(* IEC 61131-3 sources: brOscatLib/oscatBasic (part 3) *)

(* ---- REVERSE.st ---- *)
FUNCTION REVERSE
    (*http://www.oscat.de/images/OSCATBasic/oscat_basic333_en.pdf#page=232*)
    (* new code donated by rebler wolfgang *)
    REVERSE := ROR(IN,1) AND 2#10001000 OR ROL(IN,1) AND 2#00010001 OR ROR(IN,3) AND 2#01000100 OR ROL(IN,3) AND 2#00100010;

    (* old code
    REVERSE := SHL(IN,7) OR SHR(IN,7) OR (ROR(IN,3) AND 2#01000100) OR (ROL(IN,3) AND 2#00100010)
    	OR (SHL(IN,1) AND 2#00010000) OR (SHR(IN,1) AND 2#00001000);
    *)

    (* revision history
    hm		9.oct 2007		rev 1.0
    	original version

    hm		18. feb 2008	rev 1.1
    	improved performance

    RW    3. feb. 2021  	rev 1.2
    	improved performance
    *)
END_FUNCTION

(* ---- RND.st ---- *)
FUNCTION RND
    (*http://www.oscat.de/images/OSCATBasic/oscat_basic333_en.pdf#page=64*)
    IF X = 0.0 THEN
    	RND := 0.0;
    ELSE
    	M := EXPN(10.0,N - CEIL(LOG(ABS(X))));
    	RND := DINT_TO_REAL(REAL_TO_DINT(X * M)) / M;
    END_IF

    (* revision history
    hm	11. mar 2008	rev 1.0
    	original version

    hm	26. oct. 2008	rev 1.1
    	code optimization

    hm	10. mar. 2009	rev 1.2
    	real constants updated to new systax using dot

    *)

END_FUNCTION

(* ---- ROUND.st ---- *)
FUNCTION ROUND
    (*http://www.oscat.de/images/OSCATBasic/oscat_basic333_en.pdf#page=65*)
    X := cDECADES[LIMIT(0,N,8)];
    ROUND := DINT_TO_REAL(REAL_TO_DINT(IN * X)) / X;

    (* revision history
    hm	1. sep 2006	rev 1.0
    	original version

    hm	2. dec 2007	rev 1.1
    	changed code for better performance

    hm	8. jan 2008	rev 1.2
    	further improvement IN performance

    hm 11. mar. 2008	rev 1.3
    	corrected an error with negative numbers
    	use real_to_dint instead of trunc

    hm	16. mar 2008	rev 1.4
    	added type conversion to avoid warning under codesys 3.0

    hm	25. oct. 2008	rev 1.5
    	new code using global constants decades
    *)

END_FUNCTION

(* ---- SCALE.st ---- *)
FUNCTION SCALE
    (*http://www.oscat.de/images/OSCATBasic/oscat_basic333_en.pdf#page=288*)
    SCALE := LIMIT(MN, X * K + O, MX);

    (* revision history
    hm	16. may. 2008		rev 1.0
    	original version
    *)
END_FUNCTION

(* ---- SCALE_B.st ---- *)
FUNCTION SCALE_B
    (*http://www.oscat.de/images/OSCATBasic/oscat_basic333_en.pdf#page=289*)
    _I_HI := BYTE_TO_USINT(I_HI);
    _I_LO := BYTE_TO_USINT(I_LO);
    IF I_HI = I_LO THEN
    	SCALE_B := O_LO;
    ELSE
    	SCALE_B := (O_HI - O_LO) / USINT_TO_REAL(_I_HI - _I_LO) * USINT_TO_REAL(LIMIT(_I_LO, BYTE_TO_USINT(X), _I_HI));
    END_IF

    (* revision history
    hm	18. may. 2008		rev 1.0
    	original version

    hm	18. jan 2011		rev 1.1
    	avoid division by 0

    *)
END_FUNCTION

(* ---- SCALE_B2.st ---- *)
FUNCTION SCALE_B2
    (*http://www.oscat.de/images/OSCATBasic/oscat_basic333_en.pdf#page=290*)
    SCALE_B2 := 	(((IN1_MAX - IN1_MIN)* BYTE_TO_USINT(IN1) + (IN2_MAX - IN2_MIN)* BYTE_TO_USINT(IN2)) * 0.003921569 + IN1_MIN + IN2_MIN) * K + O;

    (* revision History
    hm 19.1.2007		rev 1.1
    	changed outputs to real to avoid overflow of integer
    	added offset for better cascading of scale functions
    	changed from FB to function

    hm	6. jan 2008		rev 1.2
    	improved performance

    hm	26. oct. 2008	rev 1.3
    	code optimization

    hm	3. nov. 2008	rev 1.4
    	used wrong factor in formula

    *)
END_FUNCTION

(* ---- SCALE_B4.st ---- *)
FUNCTION SCALE_B4
    (*http://www.oscat.de/images/OSCATBasic/oscat_basic333_en.pdf#page=291*)
    SCALE_B4 := 	(((IN1_MAX - IN1_MIN)* BYTE_TO_USINT(IN1) + (IN2_MAX - IN2_MIN)* BYTE_TO_USINT(IN2) + (IN3_MAX - IN3_MIN)* BYTE_TO_USINT(IN3) + (IN4_MAX - IN4_MIN)* BYTE_TO_USINT(IN4))* 0.003921569 + IN1_MIN + IN2_MIN + IN3_MIN + IN4_MIN) * K + O;

    (* revision History
    hm 19.1.2007		rev 1.1
    	changed outputs to real to avoid overflow of integer
    	added offset for better cascading of scale functions
    	changed from fb to function

    hm	6. jan 2008		rev 1.2
    	improved performance

    hm	26. oct. 2008	rev 1.3
    	optimized code

    hm	3. nov. 2008	rev 1.4
    	used wrong factor in formula

    *)
END_FUNCTION

(* ---- SCALE_B8.st ---- *)
FUNCTION SCALE_B8
    (*http://www.oscat.de/images/OSCATBasic/oscat_basic333_en.pdf#page=292*)
    SCALE_B8 := 	(((IN1_MAX - IN1_MIN)* BYTE_TO_USINT(IN1) + (IN2_MAX - IN2_MIN)* BYTE_TO_USINT(IN2) + (IN3_MAX - IN3_MIN)* BYTE_TO_USINT(IN3) + (IN4_MAX - IN4_MIN)* BYTE_TO_USINT(IN4) +
    				(IN5_MAX - IN5_MIN)* BYTE_TO_USINT(IN5) + (IN6_MAX - IN6_MIN)* BYTE_TO_USINT(IN6) + (IN7_MAX - IN7_MIN)* BYTE_TO_USINT(IN7) + (IN8_MAX - IN8_MIN)* BYTE_TO_USINT(IN8)) * 0.003921569
    				 + IN1_MIN + IN2_MIN + IN3_MIN + IN4_MIN + IN5_MIN + IN6_MIN + IN7_MIN + IN8_MIN) * K + O;

    (* revision History
    hm	19. jan.2007	rev 1.1
    	changed outputs to real to avoid overflow of integer
    	added offset for better cascading of scale functions

    hm	6. jan. 2008	rev 1.2
    	improved performance

    hm	26. oct. 2008	rev 1.3
    	code optimization

    hm	3. nov. 2008	rev 1.4
    	used wrong factor in formula

    *)
END_FUNCTION

(* ---- SCALE_D.st ---- *)
FUNCTION SCALE_D
    (*http://www.oscat.de/images/OSCATBasic/oscat_basic333_en.pdf#page=293*)
    _I_HI := DWORD_TO_UDINT(I_HI);
    _I_LO := DWORD_TO_UDINT(I_LO);
    IF _I_HI = _I_LO THEN
    	SCALE_D := O_LO;
    ELSE
    	SCALE_D := (O_HI - O_LO) / UDINT_TO_REAL(_I_HI - _I_LO) * UDINT_TO_REAL(LIMIT(_I_LO, DWORD_TO_UDINT(X), _I_HI) - _I_LO) + O_LO;
    END_IF

    (* revision history
    hm	18. may. 2008	rev 1.0
    	original version

    hm	13. nov. 2008	rev 1.1
    	corrected formula for negative gradient

    hm	11. jan 2011	rev 1.2
    	avoid division by 0
    *)
END_FUNCTION

(* ---- SCALE_R.st ---- *)
FUNCTION SCALE_R
    (*http://www.oscat.de/images/OSCATBasic/oscat_basic333_en.pdf#page=294*)
    IF I_LO = I_HI THEN
    	SCALE_R := O_LO;
    ELSE
    	SCALE_R := (O_HI - O_LO) / (I_HI - I_LO) * (LIMIT(I_LO, X, I_HI) - I_LO) + O_LO;
    END_IF

    (* revision history
    hm	18. may. 2008	rev 1.0
    	original version

    hm	13. nov. 2008	rev 1.1
    	corrected formula for negative gradient

    hm	11. jan 2011	rev 1.2
    	avoid division by 0

    *)
END_FUNCTION

(* ---- SCALE_X2.st ---- *)
FUNCTION SCALE_X2
    (*http://www.oscat.de/images/OSCATBasic/oscat_basic333_en.pdf#page=295*)
    SCALE_X2 := (SEL(IN1, IN1_MIN, IN1_MAX)+ SEL(IN2, IN2_MIN, IN2_MAX)) * K + O;

    (* revision history
    hm	19. jan, 2007	rev 1.0
    	original version

    hm	26. oct. 2008	rev 1.1
    	code optimized

    *)
END_FUNCTION

(* ---- SCALE_X4.st ---- *)
FUNCTION SCALE_X4
    (*http://www.oscat.de/images/OSCATBasic/oscat_basic333_en.pdf#page=296*)
    SCALE_X4 := (SEL(IN1,IN1_MIN, IN1_MAX) + SEL(IN2, IN2_MIN, IN2_MAX)+SEL(IN3, IN3_MIN, IN3_MAX)+ SEL(IN4, IN4_MIN, IN4_MAX)) * K + O;

    (* revision history
    hm	19. jan. 2008	rev 1.0
    	original version

    hm	26. oct. 2008	rev 1.1
    	optimized code
    *)
END_FUNCTION

(* ---- SCALE_X8.st ---- *)
FUNCTION SCALE_X8
    (*http://www.oscat.de/images/OSCATBasic/oscat_basic333_en.pdf#page=297*)
    SCALE_X8 := (SEL(IN1,IN1_MIN, IN1_MAX)+ SEL(IN2,IN2_MIN, IN2_MAX)+SEL(IN3,IN3_MIN, IN3_MAX)+ SEL(IN4,IN4_MIN, IN4_MAX)
    				+SEL(IN5,IN5_MIN, IN5_MAX)+ SEL(IN6,IN6_MIN, IN6_MAX)+SEL(IN7,IN7_MIN, IN7_MAX)+ SEL(IN8,IN8_MIN, IN8_MAX)) * K + O;

    (* revision history
    hm	19. jan. 2008	rev 1.0
    	original version

    hm	26. oct. 2008	rev 1.1
    	optimized code

    hm	24. jan. 2008	rev 1.2
    	corrected error in formula
    *)
END_FUNCTION

(* ---- SDT_TO_DATE.st ---- *)
FUNCTION SDT_TO_DATE
    (*http://www.oscat.de/images/OSCATBasic/oscat_basic333_en.pdf#page=134*)
    SDT_TO_DATE := SET_DATE(DTI.YEAR, DTI.MONTH, DTI.DAY);

    (* revision history

    hm 18. oct. 2008	rev 1.0
    	original version

    *)
END_FUNCTION

(* ---- SDT_TO_DT.st ---- *)
FUNCTION SDT_TO_DT
    (*http://www.oscat.de/images/OSCATBasic/oscat_basic333_en.pdf#page=135*)
    SDT_TO_DT := SET_DT(DTI.YEAR, DTI.MONTH, DTI.DAY, DTI.HOUR, DTI.MINUTE, DTI.SECOND);

    (* revision history

    hm 18. oct. 2008	rev 1.0
    	original version

    *)
END_FUNCTION

(* ---- SDT_TO_TOD.st ---- *)
FUNCTION SDT_TO_TOD
    (*http://www.oscat.de/images/OSCATBasic/oscat_basic333_en.pdf#page=135*)
    SDT_TO_TOD := UDINT_TO_TOD(INT_TO_UDINT(DTI.HOUR) * 3600000 + INT_TO_UDINT(DTI.MINUTE) * 60000 + INT_TO_UDINT(DTI.SECOND) * 1000 + INT_TO_UDINT(DTI.MS));

    (* revision history

    hm 18. oct. 2008	rev 1.0
    	original version

    hm	16. nov. 2008	rev 1.1
    	added typecasts to avoid warnings
    *)
END_FUNCTION

(* ---- SECOND.st ---- *)
FUNCTION SECOND
    (*http://www.oscat.de/images/OSCATBasic/oscat_basic333_en.pdf#page=135*)
    SECOND := UDINT_TO_REAL(TOD_TO_UDINT(ITOD) - TOD_TO_UDINT(ITOD)/60000 * 60000) / 1000.0;

    (* change history

    hm	2. oct. 2006 rev 1.1
    	changed name of input to ITOD

    *)
END_FUNCTION

(* ---- SECOND_OF_DT.st ---- *)
FUNCTION SECOND_OF_DT
    (*http://www.oscat.de/images/OSCATBasic/oscat_basic333_en.pdf#page=136*)
    SECOND_OF_DT := UDINT_TO_INT(DT_TO_UDINT(XDT) MOD 60);

    (* revision history
    hm		6.9.2008	rev 1.0
    	original version

    *)
END_FUNCTION

(* ---- SECOND_TO_TIME.st ---- *)
FUNCTION SECOND_TO_TIME
    (*http://www.oscat.de/images/OSCATBasic/oscat_basic333_en.pdf#page=136*)
    SECOND_TO_TIME := DWORD_TO_TIME(REAL_TO_DWORD(IN * 1000.0));

    (* revision history
    hm	4. aug. 2006	rev 1.0
    	original version

    hm	14. mar. 2008	rev 1.1
    	rounded the input after the last digit

    hm	24. feb. 2009	rev 1.2
    	changed input to IN
    *)
END_FUNCTION

(* ---- SENSOR_INT.st ---- *)
FUNCTION SENSOR_INT
    (*http://www.oscat.de/images/OSCATBasic/oscat_basic333_en.pdf#page=324*)
    IF CURRENT <> 0.0 THEN
    	RG := VOLTAGE / CURRENT;
    	SENSOR_INT := RP * ( RG - RS) / ( RP + RS - RG);
    END_IF

    (* revisaion history

    hm 20.1.2007		rev 1.1
    	deleted input R0 which was not needed.

    hm	2. dec 2007	rev 1.2
    	corrected an error in formula and improoved speed

    hm	11. mar. 2009	rev 1.3
    	changed real constants to use dot syntax

    *)
END_FUNCTION

(* ---- SET_DATE.st ---- *)
FUNCTION SET_DATE
    (*http://www.oscat.de/images/OSCATBasic/oscat_basic333_en.pdf#page=136*)
    IF (MONTH > 2) AND (SHL(YEAR,14) = 0)
    THEN (* we add one DAY for leap YEAR *)
    	SET_DATE := UDINT_TO_DATE((INT_TO_UDINT(ofs[MONTH] + DAY ) + SHR(INT_TO_UDINT(YEAR) * 1461 - 2878169, 2))*86400);
    ELSE
    	SET_DATE := UDINT_TO_DATE((INT_TO_UDINT(ofs[MONTH] + DAY - 1 ) + SHR(INT_TO_UDINT(YEAR) * 1461 - 2878169, 2))*86400);
    END_IF

    (* old code
    IF MONTH > 2 THEN
    	count := (MONTH - 1) * 30;
    	IF MONTH > 7 THEN count := count + SHR(MONTH - 3,1); ELSE count := count + SHR(MONTH - 4,1); END_IF
    	(* chech for leap YEAR and add one DAY if true
    	IF SHL(YEAR,14) = 0 THEN count := count + 1; END_IF
    ELSE
    	count := (MONTH - 1) * 31;
    END_IF

    SET_DATE := UDINT_TO_DATE((INT_TO_UDINT(count + DAY - 1) + SHR(INT_TO_UDINT(YEAR) * 1461 - 2878169, 2)) * 86400);
    *)

    (* revision history
    hm	4. aug. 2006	rev 1.0
    	original version

    hm	19 sep. 2007	rev 1.1
    	use function leap_year to calculate leap YEAR, more exceptions are handled

    hm	1. okt	2007	rev 1.2
    	added compatibility to step7

    hm	16.dec 2007		rev 1.3
    	changed code to improove performance

    hm	3. jan. 2008	rev 1.4
    	further improvements in performance

    hm	16. mar. 2008	rev 1.5
    	added type conversions to avoid warnings under codesys 3.0

    hm	7. apr. 2008	rev 1.6
    	deleted unused step7 code

    hm	14. oct. 2008	rev 1.7
    	optimized code for better performance

    hm	25. oct. 2008	rev 2.0
    	new code using setup constants

    hm	16. nov. 2008	rev 2.1
    	added typecasts to avoid warnings

    hm	22. jan. 2011	rev 2.2
    	improved performance

    hm	29. dec. 2011	rev 2.3
    	improved performance

    hm 3. FEB 2021 rev 2.4
    	new code to be more readable
    *)
END_FUNCTION

(* ---- SET_DT.st ---- *)
FUNCTION SET_DT
    (*http://www.oscat.de/images/OSCATBasic/oscat_basic333_en.pdf#page=137*)
    SET_DT := UDINT_TO_DT(DATE_TO_UDINT(SET_DATE(YEAR, MONTH, DAY)) + INT_TO_UDINT(SECOND) + INT_TO_UDINT(MINUTE) * 60 + INT_TO_UDINT(HOUR) * 3600);

    (* revision history
    hm	4. aug. 2006		rev 1.0
    	original version

    hm		19 sep. 2007	rev 1.1
    	use function leap_year to calculate leap YEAR, more exceptions are handled

    hm		1. okt 2007		rev 1.2
    	added step7 compatibility
    	call function set_date

    hm		8. oct 2007		rev 1.3
    	deleted unused variables count and leap

    hm		1. 11 2007		rev 1.4
    	converted HOUR type integer to dword in calculation to avoid overrun on möller ecp4

    hm		16. mar 2008	rev 1.5
    	added type conversions to avoid warnings under codesys 3.0
    *)

END_FUNCTION

(* ---- SET_TOD.st ---- *)
FUNCTION SET_TOD
    (*http://www.oscat.de/images/OSCATBasic/oscat_basic333_en.pdf#page=138*)
    SET_TOD := UDINT_TO_TOD(REAL_TO_UDINT(SECOND * 1000.0) + INT_TO_UDINT(MINUTE) * 60000 + INT_TO_UDINT(HOUR) * 3600000);

    (* revision history

    hm		4.aug.2006		rev 1.0
    	original version

    hm		11. sep 2007	rev 1.1
    	changed coding to avoid a compiler warning under twincat.

    hm		1. nov 2007	rev 1.2
    	changed coding to avoid possible overrun situation on möller ecp4

    hm		2. Nov	2007	rev 1.3
    	changed dword to DINT in calcualtion to avoid warnings with some compilers

    hm		14. mar 2008	rev 1.4
    	changed code to avoid rounding problem at last digit of millisecond

    hm		16. mar. 2008	rev 1.5
    	added type conversions to avoid warning under codesys 3.0
    *)
END_FUNCTION

(* ---- SGN.st ---- *)
FUNCTION SGN
    (*http://www.oscat.de/images/OSCATBasic/oscat_basic333_en.pdf#page=65*)
    IF X > 0 THEN
    	SGN := 1;
    ELSIF X < 0 THEN
    	SGN := -1;
    ELSE
    	SGN := 0;
    END_IF

    (* revision histroy
    hm	16. oct 2007	rev 1.0
    	original version

    hm	11. nov 2007	rev 1.1
    	changed type of function from real to int

    *)
END_FUNCTION

(* ---- SHL1.st ---- *)
FUNCTION SHL1
    (*http://www.oscat.de/images/OSCATBasic/oscat_basic333_en.pdf#page=233*)
    SHL1 := SHR(temp,32-N) OR SHL(IN,N);

    (* revision history
    hm	14.9.2007		rev 1.0
    	original version

    hm	27. dec 2007	rev 1.1
    	changed code for better performance

    *)
END_FUNCTION

(* ---- SHR1.st ---- *)
FUNCTION SHR1
    (*http://www.oscat.de/images/OSCATBasic/oscat_basic333_en.pdf#page=233*)
    SHR1 := SHL(temp,32-N) OR SHR(IN,N);

    (* revision history
    hm	14.9.2007		rev 1.0
    	original version

    hm	27. dec 2007	rev 1.1
    	changed code for better performance

    *)
END_FUNCTION

(* ---- SIGMOID.st ---- *)
FUNCTION SIGMOID
    (*http://www.oscat.de/images/OSCATBasic/oscat_basic333_en.pdf#page=66*)
    IF X > 20.0 THEN
    	SIGMOID := 1.0;
    ELSIF X < -85.0 THEN
    	SIGMOID := 0.0;
    ELSE
    	SIGMOID := 1.0 / (1.0 + EXP(-X));
    END_IF

    (* revision history
    hm	10.12.2007		rev 1.0
    	original version

    hm	11. mar. 2008		rev 1.1
    	extended range of valid inputs to +inv / -inv

    hm 10. mar. 2009		rev 1.2
    	real constants updated to new systax using dot

    *)
END_FUNCTION

(* ---- SIGN_I.st ---- *)
FUNCTION SIGN_I
    (*http://www.oscat.de/images/OSCATBasic/oscat_basic333_en.pdf#page=66*)
    SIGN_I := IN.31;

    (* revision history
    hm 3.3.2007	rev 1.1
    	changed method of function for better compatibility to other systems

    hm	1.12.2007	rev 1.2
    	changed code to improve performance

    hm	27. oct. 2008	rev 1.3
    	changed type of input to dint

    *)
END_FUNCTION

(* ---- SIGN_R.st ---- *)
FUNCTION SIGN_R
    (*http://www.oscat.de/images/OSCATBasic/oscat_basic333_en.pdf#page=67*)
    SIGN_R := IN < 0.0;

    (* revision history
    hm 19.1.2007	rev 1.1
    	changed method of function for better compatibility to other systems

    hm	1.12.2007	rev 1.2
    	changed code to improve performance

    hm	14. jun. 2008	rev 1.3
    	improved performace

    hm 10. mar. 2009	rev 1.4
    	real constants updated to new systax using dot

    *)
END_FUNCTION

(* ---- SINC.st ---- *)
FUNCTION SINC
    (*http://www.oscat.de/images/OSCATBasic/oscat_basic333_en.pdf#page=67*)
    IF X = 0.0 THEN
    	SINC := 1.0;
    ELSE
    	SINC := SIN(X) / X;
    END_IF

    (* revision histroy
    hm	11. mar. 2008	rev 1.0
    	original version

    hm	1.12.2007	rev 1.1
    	changed code to improove performance

    hm 10. mar. 2009	rev 1.2
    	real constants updated to new systax using dot

    *)
END_FUNCTION

(* ---- SINH.st ---- *)
FUNCTION SINH
    (*http://www.oscat.de/images/OSCATBasic/oscat_basic333_en.pdf#page=67*)
    IF ABS(X) < 2E-3 THEN
    	SINH := X;
    ELSE
    	SINH := (EXP(X) - EXP(-X)) * 0.5;
    END_IF

    (* revision history
    hm	12.1.2007	rev 1.0
    	original version

    hm	1.12.2007	rev 1.1
    	changed code to improve performance

    hm	5. jan 2008	rev 1.2
    	further performance improvement

    hm	11. mar 2008	rev 1.3
    	improved accuracy around 0

    *)
END_FUNCTION

(* ---- SPHERE_V.st ---- *)
FUNCTION SPHERE_V
    (*http://www.oscat.de/images/OSCATBasic/oscat_basic333_en.pdf#page=106*)
    SPHERE_V := 4.188790205 * RX * RX * RX;

    (* revision histroy
    hm	16. oct 2007	rev 1.0
    	original version

    hm	4. dec 2007		rev 1.1
    	changed code for better performance

    hm	22. feb 2008		rev 1.2
    	changed code for better performance
    *)

END_FUNCTION

(* ---- SQRTN.st ---- *)
FUNCTION SQRTN
    (*http://www.oscat.de/images/OSCATBasic/oscat_basic333_en.pdf#page=68*)
    IF N > 0 THEN
    	SQRTN := EXP(LN(X) / INT_TO_REAL(N));
    ELSE
    	SQRTN := 0.0;
    END_IF

    (* revision history
    hm		12 jan 2007	rev 1.0
    	original version

    hm		2. dec 2007	rev 1.1
    	changed code for better performance

    hm		11. mar 2008	rev 1.2
    	added result 0 for compatibility reasons

    hm 10. mar. 2009	rev 1.3
    	added type conversions for compatibility reasons

    *)
END_FUNCTION

(* ---- STAIR.st ---- *)
FUNCTION STAIR
    (*http://www.oscat.de/images/OSCATBasic/oscat_basic333_en.pdf#page=304*)
    IF D > 0.0 THEN
    	STAIR := DINT_TO_REAL(REAL_TO_DINT(X / D)) * D;
    ELSE
    	STAIR := X;
    END_IF

    (* revision history
    hm	28 jan 2007		rev 1.0
    	original version

    hm	27 dec 2007		rev 1.1
    	changed code for better performance

    hm	6. jan 2008		rev 1.2
    	further performance improvement

    hm	26. oct. 2008		rev 1.3
    	optimized code

    hm	10. mar. 2009	rev 1.4
    	real constants updated to new systax using dot

    *)
END_FUNCTION

(* ---- STATUS_TO_ESR.st ---- *)
FUNCTION STATUS_TO_ESR
    (*http://www.oscat.de/images/OSCATBasic/oscat_basic333_en.pdf#page=38*)
    IF STATUS < 100 THEN
    	RETVAL.TYP := 1;
    ELSIF STATUS < 200 THEN
    	RETVAL.TYP := 2;
    ELSE
    	RETVAL.TYP := 3;
    END_IF
    RETVAL.ADRESS:= ADRESS;
    RETVAL.DS := DT_IN;
    RETVAL.TS := TS;
    RETVAL.DATA[0] := STATUS;
    STATUS_TO_ESR:=TRUE;
END_FUNCTION

(* ---- SUN_MIDDAY.st ---- *)
FUNCTION SUN_MIDDAY
    (*http://www.oscat.de/images/OSCATBasic/oscat_basic333_en.pdf#page=138*)
    T := INT_TO_REAL(DAY_OF_YEAR(UTC));
    OFFSET := -0.1752 * SIN(0.033430 * T + 0.5474) - 0.1340 * SIN(0.018234 * T - 0.1939);
    SUN_MIDDAY := HOUR_TO_TOD(12.0 - OFFSET - LON * 0.0666666666666);

    (* revision history

    hm	26. jan. 2011	rev 1.0
    	initial release

    *)
END_FUNCTION

(* ---- SWAP_BYTE.st ---- *)
FUNCTION SWAP_BYTE
    (*http://www.oscat.de/images/OSCATBasic/oscat_basic333_en.pdf#page=234*)
    SWAP_BYTE := ROL(IN,8);

    (* revision history
    hm		4. feb 2008	rev 1.0
    	original version

    *)
END_FUNCTION

(* ---- SWAP_BYTE2.st ---- *)
FUNCTION SWAP_BYTE2
    (*http://www.oscat.de/images/OSCATBasic/oscat_basic333_en.pdf#page=234*)
    SWAP_BYTE2 := (ROR(IN,8) AND 16#FF00FF00) OR (ROL(IN,8) AND 16#00FF00FF);

    (* revision history
    hm		4. feb 2008	rev 1.0
    	original version

    *)

END_FUNCTION

(* ---- T_PLC_MS.st ---- *)
FUNCTION T_PLC_MS
    (*http://www.oscat.de/images/OSCATBasic/oscat_basic333_en.pdf#page=348*)
    tx := TIME();
    T_PLC_MS := TIME_TO_UDINT(tx);
    (* hier muss die korrektur für step7 stattfinden
    plctime muss den vollen wertebereich von time ausnutzen:
    wenn bei step7 time -24tage bis plus 24 tage ist dann muss der timer auch beim überlauf auf -24tage springen
    und auf keinen fall auf 0 !!!!
    für siemens muss ein weiterer fb im main eingebunden werden der sicherstellt das alle 32 bits durchgezählt werden.
    es kann nur ein fb sein den er muss sich das oberste (32te) bit merken.
    oder etwa spring s7 bei überlauf auf -24 tage????? dann wäre keine korrektur nötig.
    *)
    IF debug THEN
    	T_PLC_MS := (SHL(T_PLC_MS,N) OR SHL(UDINT#1,N)-1) + offset;
    END_IF

    (* revision history
    hm	14.9.2007	rev 1.0
    	original version

    hm	12. nov 2007	rev 1.1
    	added temporaray variable tx because some compilers could not handle time() as an argument

    hm	16. nov. 2008	rev 1.2
    	initialized constants with 0 for compatibility reasons
    *)
END_FUNCTION

(* ---- T_PLC_US.st ---- *)
FUNCTION T_PLC_US
    (*http://www.oscat.de/images/OSCATBasic/oscat_basic333_en.pdf#page=351*)
    tx := TIME();
    T_PLC_US := TIME_TO_UDINT(tx)*1000;
    (* hier muss die korrektur für step7 stattfinden
    plctime muss den vollen wertebereich von time ausnutzen:
    wenn bei step7 time -24tage bis plus 24 tage ist dann muss der timer auch beim überlauf auf -24tage springen
    und auf keinen fall auf 0 !!!!
    für siemens muss ein weiterer fb im main eingebunden werden der sicherstellt das alle 32 bits durchgezählt werden.
    es kann nur ein fb sein den er muss sich das oberste (32te) bit merken.
    oder etwa spring s7 bei überlauf auf -24 tage????? dann wäre keine korrektur nötig.
    *)
    IF debug THEN
    	T_PLC_US := (SHL(T_PLC_US,N) OR SHL(UDINT#1,N)-1) + offset;
    END_IF

    (* revision history
    hm	14.9.2007	rev 1.0
    	original version

    hm	12. nov 2007	rev 1.1
    	added temporaray variable tx because some compilers could not handle time() as an argument

    hm	16. nov. 2008	rev 1.2
    	initialized constants with 0 for compatibility reasons

    *)
END_FUNCTION

(* ---- TANC.st ---- *)
FUNCTION TANC
    (*http://www.oscat.de/images/OSCATBasic/oscat_basic333_en.pdf#page=68*)
    IF X = 0.0 THEN
    	TANC := 1.0;
    ELSE
    	TANC := TAN(X) / X;
    END_IF

    (* revision histroy
    hm	23. oct. 2008	rev 1.0
    	original version

    hm 10. mar. 2009	rev 1.1
    	real constants updated to new systax using dot

    *)
END_FUNCTION

(* ---- TANH.st ---- *)
FUNCTION TANH
    (*http://www.oscat.de/images/OSCATBasic/oscat_basic333_en.pdf#page=69*)
    IF X > 20.0 THEN
    	TANH := 1.0;
    ELSIF X < -20.0 THEN
    	TANH := -1.0;
    ELSE
    	TANH := 1.0 - 2.0 / (EXP(2.0 * X) + 1.0);
    END_IF

    (* revision hisdtory
    hm		12.1.2007		rev 1.0
    	original version

    hm		1.12.2007		rev 1.1
    	changed code to improve performance

    hm		10. mar 2008	rev 1.2
    	corrected an error in formula
    	extended range of valid inputs to +/- INV

    hm 10. mar. 2009	rev 1.3
    	real constants updated to new systax using dot

    *)
END_FUNCTION

(* ---- TEMP_NI.st ---- *)
FUNCTION TEMP_NI
    (*http://www.oscat.de/images/OSCATBasic/oscat_basic333_en.pdf#page=325*)
    TEMP_NI := (SQRT(0.30085225 - 2.66E-3 * (R0 - RES)) - 0.5485) * 751.8796992;

    (* revision history

    hm 24.1.2007		rev 1.1
    	deleted unused variable A, B, C

    hm 10.9.2007		rev 1.2
    	changed accuracy to 0.02 degrees to improove performace

    hm 17. 12 2007	rev 1.3
    	improovements for better performance and higher accuracy

    hm	6. jan 2008	rev 1.4
    	further performance improvement

    hm	10. mar. 2009	rev 1.5
    	removed nested comments

    *)

END_FUNCTION

(* ---- TEMP_NTC.st ---- *)
FUNCTION TEMP_NTC
    (*http://www.oscat.de/images/OSCATBasic/oscat_basic333_en.pdf#page=326*)
    IF RES > 0.0 THEN
    	TEMP_NTC := B * 298.15 / (B + LN(RES / RN) * 298.15) -273.15;
    END_IF

    (* revision history

    hm 30. dec. 2008	rev 1.0
    	original version

    hm	11. mar. 2009	rev 1.1
    	changed real constants to use dot syntax

    *)
END_FUNCTION

(* ---- TEMP_PT.st ---- *)
FUNCTION TEMP_PT
    (*http://www.oscat.de/images/OSCATBasic/oscat_basic333_en.pdf#page=326*)
    X := A * R0;
    Y := B * R0;
    IF RES >= R0 THEN
    	t1 := X * X - 4.0 * Y * (R0 - RES);
    	IF t1 < 0.0 THEN
    		TEMP_PT := 10000.0;
    	ELSE
    		TEMP_PT := (-X + SQRT(t1)) / (2.0 * Y);
    	END_IF
    ELSE
    	pt ACCESS ADR(step);
    	(* since the formula cannot be solved this is A successive approximation *)
    	TEMP_PT := -100.0;
    	WHILE step > accuracy DO
    		(* test if result greater or less *)
    		IF RES_PT(TEMP_PT, R0) < RES THEN TEMP_PT := TEMP_PT + step; ELSE TEMP_PT := TEMP_PT - step; END_IF
    		pt := pt - 8388608;  (* this is A super fast divide by 2 method for non floating point CPUs *)
    		(* the alternative code: step := step * 0.5; *)
    	END_WHILE
    END_IF

    (* revision history

    rev 1.1 hm 24.1.2007
    	deleted unused variable C

    rev 1.2 hm 10.9.2007
    	reduced accuracy to 0.02 to shorten execution time

    rev 1.3	hm	2. dec 2007
    	changed code for better performance

    rev	1.4	hm	23. dec 2007
    	avoid A negative square root if input values are wrong

    rev 1.5 hm	5. jan 2008
    	replaced / 2 with * 0.5 for better performance

    hm	31. oct. 2008	rev 1.6
    	improved performance

    hm	11. mar. 2009	rev 1.7
    	changed real constants to use dot syntax

    *)

END_FUNCTION

(* ---- TEMP_SI.st ---- *)
FUNCTION TEMP_SI
    (*http://www.oscat.de/images/OSCATBasic/oscat_basic333_en.pdf#page=331*)
    TEMP_SI := (-7.64E-3 + SQRT(RES / RS * 6.64E-5 - 0.803E-5)) * 30120.48193 + TS;

    (* revision history

    hm 24.1.2007		rev 1.1
    	the function would only work for TS = 25, now it works for other values of TS.

    hm 10.9.2007		rev 1.2
    	changed the function to use successive approcimation to avoid an error generated by a sqrt from a negative result.
    	changed accuracy to 0.02 degrees to shorten execution time

    hm 17. 12 2007	rev 1.3
    	improovements for better performance

    hm	6. jan 2008	rev 1.4
    	further performance improvement

    hm	10. mar. 2009	rev 1.5
    	removed nested comments

    *)
END_FUNCTION

(* ---- TIMECHECK.st ---- *)
FUNCTION TIMECHECK
    (*http://www.oscat.de/images/OSCATBasic/oscat_basic333_en.pdf#page=141*)
    IF STOP < START THEN
    	TIMECHECK := START <= TD OR TD < STOP;
    ELSE
    	TIMECHECK := START <= TD AND TD < STOP;
    END_IF

    (* revision history
    hm 19. jul. 2009	rev 1.0
    	original release

    *)
END_FUNCTION

(* ---- TO_LOWER.st ---- *)
FUNCTION TO_LOWER
    (*http://www.oscat.de/images/OSCATBasic/oscat_basic333_en.pdf#page=179*)
    byteAsInt := BYTE_TO_USINT(IN);
    IF byteAsInt > 64 AND byteAsInt < 91 THEN
       TO_LOWER := IN OR 16#20;
    ELSIF (byteAsInt > 191 AND byteAsInt < 223) AND byteAsInt <> 215 AND cEXTENDED_ASCII THEN
       TO_LOWER := IN OR 16#20;
    ELSE
       TO_LOWER := IN;
    END_IF

    (* revision history
    hm	6. mar. 2008	rev 1.0
    	original version

    hm	19. oct. 2008	rev 1.1
    	changed setup constants

    ks	25. oct. 2008	rev 1.2
    	optimized code
    *)
END_FUNCTION

(* ---- TO_UML.st ---- *)
FUNCTION TO_UML
    (*http://www.oscat.de/images/OSCATBasic/oscat_basic333_en.pdf#page=180*)
    CASE BYTE_TO_USINT(IN) OF
    	196:	(* Ä *)
    		RETVAL := 'Ae';
    	214:	(* Ö *)
    		RETVAL := 'Oe';
    	220:	(* Ü *)
    		RETVAL := 'Ue';
    	223:	(* ß *)
    		RETVAL := 'ss';
    	228:	(* ä *)
    		RETVAL := 'ae';
    	246:	(* ö *)
    		RETVAL := 'oe';
    	252:	(* ü *)
    		RETVAL := 'ue';
    ELSE
    	CHR_TO_STRING(IN, RETVAL);
    END_CASE
    TO_UML := TRUE;

    (* revision history
    hm	29. mar. 2008	rev 1.0
    	original version

    hm	17. dec. 2008	rev 1.1
    	changes name of function chr to chr_to_string

    *)
END_FUNCTION

(* ---- TO_UPPER.st ---- *)
FUNCTION TO_UPPER
    (*http://www.oscat.de/images/OSCATBasic/oscat_basic333_en.pdf#page=180*)
    byteAsInt := BYTE_TO_USINT(IN);
    IF byteAsInt > 96 AND byteAsInt < 123 THEN
       TO_UPPER := IN AND 16#DF;
    ELSIF byteAsInt > 223 AND byteAsInt <> 247 AND byteAsInt <> 255 AND cEXTENDED_ASCII THEN
       TO_UPPER := IN AND 16#DF;
    ELSE
       TO_UPPER := IN;
    END_IF

    (* revision history
    hm	6. mar. 2008	rev 1.0
    	original version

    hm	19. oct. 2008	rev 1.1
    	changed setup constants

    ks	25. oct. 2008	rev 1.2
    	optimized code

    hm 16. jan 2009	rev 1.3
    	corrected an error IN module

    *)
END_FUNCTION

(* ---- TRIANGLE_A.st ---- *)
FUNCTION TRIANGLE_A
    (*http://www.oscat.de/images/OSCATBasic/oscat_basic333_en.pdf#page=107*)
    IF A = 0.0 THEN
    	TRIANGLE_A := SQRT((S1+S2+S3) * (S1+S2-S3) * (S2+S3-S1) * (S3+S1-S2)) * 0.25;
    ELSE
    	TRIANGLE_A := S1 * S2 * SIN(RAD(A)) * 0.5;
    END_IF

    (* revision histroy
    hm	16. oct 2007	rev 1.0
    	original version

    hm	22. feb 2008	rev 1.1
    	improved performance

    hm	10. mar. 2009	rev 1.2
    	changed syntax of real constants to 0.0

    *)
END_FUNCTION

(* ---- TRIM.st ---- *)
FUNCTION TRIM
    (*http://www.oscat.de/images/OSCATBasic/oscat_basic333_en.pdf#page=181*)
    RETVAL := STR;
    REPEAT
    	pos := FIND(RETVAL,' ');
    	IF pos > 0 THEN RETVAL := REPLACE(RETVAL,'',1,pos); END_IF
    UNTIL pos = 0	END_REPEAT
    TRIM := TRUE;

    (* revision histroy
    hm	6.10.2006		rev 1.0
    	original release

    hm	20. mar. 2008	rev 1.1
    	avoid to call replace with pos = 0 because some systems will produce an error

    hm	29. mar. 2008	rev 1.2
    	changed STRING to STRING(STRING_LENGTH)
    *)
END_FUNCTION

(* ---- TRIM1.st ---- *)
FUNCTION TRIM1
    (*http://www.oscat.de/images/OSCATBasic/oscat_basic333_en.pdf#page=181*)
    RETVAL := STR;
    REPEAT
    	pos := FIND(RETVAL,'  ');
    	IF pos > 0 THEN RETVAL := REPLACE(RETVAL,' ',2,pos); END_IF
    UNTIL pos = 0	END_REPEAT
    (* beginning and ending blanks need to be stripped off *)
    IF LEFT(RETVAL,1) = ' ' THEN RETVAL := DELETE(RETVAL,1,1); END_IF
    IF RIGHT(RETVAL,1) = ' ' THEN RETVAL := DELETE(RETVAL,1,LEN(RETVAL)); END_IF
    TRIM1 := TRUE;

    (* revision histroy
    hm	4. feb. 2008    rev 1.0
    	original release

    hm	20. mar. 2008	rev 1.1
    	avoid to call replace with pos = 0 because some systems will produce an error

    hm	29. mar. 2008	rev 1.2
    	changed STRING to STRING(STRING_LENGTH)
    *)
END_FUNCTION

(* ---- TRIME.st ---- *)
FUNCTION TRIME
    (*http://www.oscat.de/images/OSCATBasic/oscat_basic333_en.pdf#page=181*)
    RETVAL := STR;
    (* beginning blanks need to be stripped off *)
    WHILE LEFT(RETVAL,1) = ' ' DO
    	RETVAL := DELETE(RETVAL,1,1);
    END_WHILE

    (* ending blanks need to be stripped off *)
    WHILE RIGHT(RETVAL,1) = ' ' DO
    	RETVAL := DELETE(RETVAL,1,LEN(RETVAL));
    END_WHILE
    TRIME := TRUE;

    (* revision histroy
    hm	28. mar. 2008	rev 1.0
    	original release

    *)
END_FUNCTION

(* ---- UPPERCASE.st ---- *)
FUNCTION UPPERCASE
    (*http://www.oscat.de/images/OSCATBasic/oscat_basic333_en.pdf#page=182*)
    pt ACCESS ADR(RETVAL);
    RETVAL := STR;
    l := LEN(STR);
    FOR pos := 1 TO l DO
    	pt := TO_UPPER(pt);
    	pt ACCESS (ADR(pt) + 1);
    END_FOR
    UPPERCASE := TRUE;

    (* revision histroy
    hm	6. oct. 2006	rev 1.0
    	original release

    hm	4. feb. 2008	rev 1.1
    	improved performance
    	added Ä,Ö,Ü

    hm	6. mar. 2008	rev 1.2
    	added support for exteded Ascii

    hm	29. mar. 2008	rev 1.3
    	changed STRING to STRING(STRING_LENGTH)

    *)

END_FUNCTION

(* ---- UTC_TO_LTIME.st ---- *)
FUNCTION UTC_TO_LTIME
    (*http://www.oscat.de/images/OSCATBasic/oscat_basic333_en.pdf#page=142*)
    tmp := TIME_ZONE_OFFSET * 60 + BOOL_TO_INT(DST_ENABLE AND DST(UTC)) * 3600;
    IF tmp < 0 THEN
    	tmp := ABS(tmp);
    	UTC_TO_LTIME := UDINT_TO_DT(DT_TO_UDINT(UTC) -  INT_TO_UDINT(tmp));
    ELSE
    	UTC_TO_LTIME := UDINT_TO_DT(DT_TO_UDINT(UTC) +  INT_TO_UDINT(tmp));
    END_IF

    (* revision history

    hm 2.10.2006	rev 1.1
    	corrected an error where dst would be delayed by 0.1second

    hm 17.1.2007	rev 1.2
    	added UTC input instead of internal sysrtcgettime because this would only work on wago.
    	DST_ENABLE would not be checked before dst would be enabled.

    hm 18.3.2007	rev 1.3
    	changed code, dst would not work during first cycle.

    hm 24.10.2007	rev 1.4
    	changed code because the execution every 100ms can cause major problems if the supplied time was not correct at start.
    	use of new dst function

    hm 12. nov 2007	rev 1.5
    		changed Type of TIME_ZONE_OFFSET from time to int to allow for time zones with negative offset

    hm	8 dec 2007		rev 1.6
    	corrected a problem with TIME_ZONE_OFFSET

    hm	14. oct. 2008	rev 1.7
    	renamed module from LTIME to UTC_TO_LTIME
    	changed function weekday to day_of_week
    	optimized code for better performance

    hm	20. oct. 2008	rev 1.8
    	changes type of input TIME_ZONE_OFFSET from real to int, now is in +/-minutes
    	deleted outputs DST_ON and WDAY
    	converted to function

    hm	27. feb. 2009	rev 1.9
    	added type conversions to avoid warnings under codesys 3.0

    *)
END_FUNCTION

(* ---- V3_ABS.st ---- *)
FUNCTION V3_ABS
    (*http://www.oscat.de/images/OSCATBasic/oscat_basic333_en.pdf#page=108*)
    V3_ABS := SQRT(A.X * A.X + A.Y * A.Y + A.Z * A.Z);

    (* revision history
    hm		11 dec 2007	rev 1.0
    	original version

    *)
END_FUNCTION

(* ---- V3_ADD.st ---- *)
FUNCTION V3_ADD
    (*http://www.oscat.de/images/OSCATBasic/oscat_basic333_en.pdf#page=108*)
    RETVAL.X := A.X + B.X;
    RETVAL.Y := A.Y + B.Y;
    RETVAL.Z := A.Z + B.Z;
    V3_ADD:=TRUE;

    (* revision history
    hm		11 dec 2007	rev 1.0
    	original version

    *)
END_FUNCTION

(* ---- V3_ANG.st ---- *)
FUNCTION V3_ANG
    (*http://www.oscat.de/images/OSCATBasic/oscat_basic333_en.pdf#page=109*)
    d := V3_ABS(A) * V3_ABS(B);
    IF d > 0 THEN
    	V3_ANG := ACOS(LIMIT(-1.0, V3_DPRO(A, B) / d,1.0));
    END_IF

    (* revision history
    hm	11. dec. 2007	rev 1.0
    	original version

    hm	10. mar. 2009	rev 1.1
    	changed syntax of real constants to 0.0

    *)
END_FUNCTION

(* ---- V3_DPRO.st ---- *)
FUNCTION V3_DPRO
    (*http://www.oscat.de/images/OSCATBasic/oscat_basic333_en.pdf#page=109*)
    V3_DPRO := A.X * B.X + A.Y * B.Y + A.Z * B.Z;

    (* revision history
    hm		11 dec 2007	rev 1.0
    	original version

    *)
END_FUNCTION

(* ---- V3_NORM.st ---- *)
FUNCTION V3_NORM
    (*http://www.oscat.de/images/OSCATBasic/oscat_basic333_en.pdf#page=110*)
    la := V3_ABS(A);
    IF la > 0.0 THEN
    	V3_SMUL(A, 1.0 / la, RETVAL);
        V3_NORM := TRUE;
    ELSE
        V3_NORM := FALSE;
    END_IF

    (* revision history
    hm	11 dec 2007	rev 1.0
    	original version

    hm	10. mar. 2009	rev 1.1
    	changed syntax of real constants to 0.0

    *)
END_FUNCTION

(* ---- V3_NUL.st ---- *)
FUNCTION V3_NUL
    (*http://www.oscat.de/images/OSCATBasic/oscat_basic333_en.pdf#page=110*)
    V3_NUL := A.X = 0.0 AND A.Y = 0.0 AND A.Z = 0.0;

    (* revision history
    hm	12 dec 2007	rev 1.0
    	original version

    hm	10. mar. 2009	rev 1.1
    	changed syntax of real constants to 0.0

    *)
END_FUNCTION

(* ---- V3_PAR.st ---- *)
FUNCTION V3_PAR
    (*http://www.oscat.de/images/OSCATBasic/oscat_basic333_en.pdf#page=110*)
    V3_XPRO(A, B,temp);
    V3_PAR := V3_ABS(temp) = 0.0;

    (* revision history
    hm	11 dec 2007	rev 1.0
    	original version

    hm	10. mar. 2009	rev 1.1
    	changed syntax of real constants to 0.0

    *)
END_FUNCTION

(* ---- V3_REV.st ---- *)
FUNCTION V3_REV
    (*http://www.oscat.de/images/OSCATBasic/oscat_basic333_en.pdf#page=111*)
    RETVAL.X := -A.X;
    RETVAL.Y := -A.Y;
    RETVAL.Z := -A.Z;
    V3_REV:=TRUE;

    (* revision history
    hm		11 dec 2007	rev 1.0
    	original version

    *)
END_FUNCTION

(* ---- V3_SMUL.st ---- *)
FUNCTION V3_SMUL
    (*http://www.oscat.de/images/OSCATBasic/oscat_basic333_en.pdf#page=111*)
    RETVAL.X := A.X * M;
    RETVAL.Y := A.Y * M;
    RETVAL.Z := A.Z * M;
    V3_SMUL:=TRUE;

    (* revision history
    hm		11 dec 2007	rev 1.0
    	original version

    *)
END_FUNCTION

(* ---- V3_SUB.st ---- *)
FUNCTION V3_SUB
    (*http://www.oscat.de/images/OSCATBasic/oscat_basic333_en.pdf#page=112*)
    RETVAL.X := A.X - B.X;
    RETVAL.Y := A.Y - B.Y;
    RETVAL.Z := A.Z - B.Z;
    V3_SUB := TRUE;

    (* revision history
    hm		11 dec 2007	rev 1.0
    	original version

    *)
END_FUNCTION

(* ---- V3_XANG.st ---- *)
FUNCTION V3_XANG
    (*http://www.oscat.de/images/OSCATBasic/oscat_basic333_en.pdf#page=112*)
    la := V3_ABS(A);
    IF la > 0.0 THEN
    	V3_XANG := ACOS(A.X / la);
    END_IF

    (* revision history
    hm	11 dec 2007	rev 1.0
    	original version

    hm	10. mar. 2009	rev 1.1
    	changed syntax of real constants to 0.0

    *)
END_FUNCTION

(* ---- V3_XPRO.st ---- *)
FUNCTION V3_XPRO
    (*http://www.oscat.de/images/OSCATBasic/oscat_basic333_en.pdf#page=112*)
    RETVAL.X := A.Y * B.Z - A.Z * B.Y;
    RETVAL.Y := A.Z * B.X - A.X * B.Z;
    RETVAL.Z := A.X * B.Y - A.Y * B.X;
    V3_XPRO:=TRUE;

    (* revision history
    hm		11 dec 2007	rev 1.0
    	original version

    *)
END_FUNCTION

(* ---- V3_YANG.st ---- *)
FUNCTION V3_YANG
    (*http://www.oscat.de/images/OSCATBasic/oscat_basic333_en.pdf#page=113*)
    la := V3_ABS(A);
    IF la > 0.0 THEN
    	V3_YANG := ACOS(A.Y / la);
    END_IF

    (* revision history
    hm	11 dec 2007	rev 1.0
    	original version

    hm	10. mar. 2009	rev 1.1
    	changed syntax of real constants to 0.0

    *)
END_FUNCTION

(* ---- V3_ZANG.st ---- *)
FUNCTION V3_ZANG
    (*http://www.oscat.de/images/OSCATBasic/oscat_basic333_en.pdf#page=113*)
    la := V3_ABS(A);
    IF la > 0.0 THEN
    	V3_ZANG := ACOS(A.Z / la);
    END_IF

    (* revision history
    hm	11 dec 2007	rev 1.0
    	original version

    hm	10. mar. 2009	rev 1.1
    	changed syntax of real constants to 0.0

    *)
END_FUNCTION

(* ---- WEEKDAY_TO_STRING.st ---- *)
FUNCTION WEEKDAY_TO_STRING
    (*http://www.oscat.de/images/OSCATBasic/oscat_basic333_en.pdf#page=182*)
    IF LANG = 0 THEN ly := cLANGUAGE_DEFAULT; ELSE ly := MIN(LANG, cLANGUAGE_LMAX); END_IF
    IF WDAY < 1 OR WDAY > 7 THEN
    	RETURN;
    ELSIF LX = 0 THEN
    	RETVAL := cWEEKDAYS[ly, WDAY];
    ELSIF LX = 2 THEN
    	RETVAL := cWEEKDAYS2[ly, WDAY];
    END_IF
    WEEKDAY_TO_STRING := TRUE;

    (* revisison history

    hm	21. sep. 2008	rev 1.0
    	original version

    hm	19. oct. 2008	rev 1.1
    	changed language setup constants
    *)
END_FUNCTION

(* ---- WINDOW.st ---- *)
FUNCTION WINDOW
    (*http://www.oscat.de/images/OSCATBasic/oscat_basic333_en.pdf#page=69*)
    WINDOW := IN < HIGH AND IN > LOW;

    (* revision history
    hm	22.1.2007	rev 1.1
    	changed the order of inputs to LOW, IN, HIGH

    *)
END_FUNCTION

(* ---- WINDOW2.st ---- *)
FUNCTION WINDOW2
    (*http://www.oscat.de/images/OSCATBasic/oscat_basic333_en.pdf#page=69*)
    WINDOW2 := IN >= LOW AND IN <= HIGH;

    (* revision history
    hm	31.10.2007	rev 1.0
    	original version

    *)
END_FUNCTION

(* ---- WORD_OF_BYTE.st ---- *)
FUNCTION WORD_OF_BYTE
    (*http://www.oscat.de/images/OSCATBasic/oscat_basic333_en.pdf#page=234*)
    WORD_OF_BYTE := SHL(BYTE_TO_WORD(B1),8) OR BYTE_TO_WORD(B0);

    (* revision history
    hm	24. jan 2007	rev 1.0
    	original version

    hm	2. jan 2008	rev 1.1
    	improved performance

    hm	19. feb 2008	rev 1.2
    	replaced and with or for better compatibility

    hm	23. apr. 2008	rev 1.3
    	reverse order of inputs to be more logical

    hm	18. jul. 2009	rev 1.4
    	added type conversions for compatibility reasons

    *)
END_FUNCTION

(* ---- WORD_OF_DWORD.st ---- *)
FUNCTION WORD_OF_DWORD
    (*http://www.oscat.de/images/OSCATBasic/oscat_basic333_en.pdf#page=235*)
    WORD_OF_DWORD := DWORD_TO_WORD(SHR(IN,SHL(N,4)));

    (* revision history
    hm	17. jan 2007	rev 1.0
    	original version

    hm	2. jan 2008		rev 1.1
    	improved performance

    hm	30. oct. 2008	rev 1.2
    	improved performance
    *)

END_FUNCTION

(* ---- WORD_TO_RANGE.st ---- *)
FUNCTION WORD_TO_RANGE
    (*http://www.oscat.de/images/OSCATBasic/oscat_basic333_en.pdf#page=316*)
    WORD_TO_RANGE := (HIGH - LOW) * WORD_TO_REAL(X) * 0.00001525902189669640 + LOW;

    (* revision history
    hm	9. jan 2008	rev 1.0
    	original version

    hm	10. mar. 2009	rev 1.1
    	improved code
    *)

END_FUNCTION

(* ---- WORK_WEEK.st ---- *)
FUNCTION WORK_WEEK
    (*http://www.oscat.de/images/OSCATBasic/oscat_basic333_en.pdf#page=142*)
    (* berechne den 1.1 des jahres von IDATE. *)
    yr := YEAR_OF_DATE(IDATE);
    d1 := YEAR_BEGIN(yr);
    (* wochentag von d1 *)
    w1 := DAY_OF_WEEK(d1);
    (* offset des montags der eletzten KW des vorjahres *)
    (* wenn der erste tag des jahres größer als donnerstag ist dann beginnt die letzte kw am montag davor *)
    (* wenn der erste tag des jahres ein donnerstag oder kleiner ist beginnt die erste kw 2 montage davor *)
    IF w1 < 5 THEN
    	ds := DATE_TO_UDINT(d1) - INT_TO_UDINT(w1+6) * 86400;
    ELSE
    	ds := DATE_TO_UDINT(d1) - INT_TO_UDINT(w1-1) * 86400;
    END_IF

    (* kalenderwoche des eingangsdatums *)
    WORK_WEEK := UDINT_TO_INT((DATE_TO_UDINT(IDATE) - ds) / 604800);

    (* korrektur wenn WORK_WEEK = 0 *)
    IF WORK_WEEK = 0 THEN
    	(* WORK_WEEK needs to be 53 when 1.jan of the year before is thursday or dec 31. is thursday. *)
    	(* first and last weekday of a year is equal and one more day for a LEAP_YEAR. *)
    	IF w1 > 1 THEN w31 := w1 - 1; ELSE w31 := 7; END_IF
    	IF LEAP_YEAR(yr - 1) AND w31 > 1 THEN w01 := w31 - 1; ELSE w1 := 7; END_IF
    	(* if first or last day of a year is a thursday, the year has 53 weeks *)
    	WORK_WEEK := 52 + BOOL_TO_INT(w31 = 4 OR w01 = 4);
    ELSE
    	(* end of year calculation *)
    	(* calculated the first and last weekday *)
    	IF LEAP_YEAR(yr) THEN
    		IF w1 < 7 THEN w31 := w1 + 1; ELSE w31 := 1; END_IF
    	ELSE
    		w31 := w1;
    	END_IF
    	(* if first or last day is thursday then the year has 53 weeks otherwise only 52 *)
    	wm := 52 + BOOL_TO_INT(w31 = 4 OR w1 = 4);
    	IF WORK_WEEK > wm THEN WORK_WEEK := 1; END_IF
    END_IF

    (* revision history

    hm 	17.1.2007		rev 1.1
    	deleted unused variable yday

    hm	19. dec 2007	rev 1.2
    	changed code for better performance
    	changed code to comply with ISO8601

    hm	16. mar 2008	rev 1.3
    	added type conversions to avoid warnings under codesys 3.0

    hm	7. oct. 2008	rev 1.4
    	changed function year to year_of_date
    	changed function weekday to day_of_week

    hm	25. oct. 2008	rev 1.5
    	optimized code for performance
    *)
END_FUNCTION

(* ---- YEAR_BEGIN.st ---- *)
FUNCTION YEAR_BEGIN
    (*http://www.oscat.de/images/OSCATBasic/oscat_basic333_en.pdf#page=143*)
    YEAR_BEGIN := UDINT_TO_DATE(SHR(INT_TO_UDINT(Y) * 1461 - 2878169,2) * 86400);

    (* revision history
    hm	19. dec 2007	rev 1.0
    	original version

    hm	4. jan 2008		rev 1.1
    	formula for step7 was incorrect during leap years

    hm	7. apr. 2008	rev 1.2
    	deleted unused step7 code
    *)

END_FUNCTION

(* ---- YEAR_END.st ---- *)
FUNCTION YEAR_END
    (*http://www.oscat.de/images/OSCATBasic/oscat_basic333_en.pdf#page=143*)
    YEAR_END := UDINT_TO_DATE(SHR(INT_TO_UDINT(Y) * 1461 - 2876712, 2) * 86400);

    (* revision history
    hm	15. jun. 2008	rev 1.0
    	original version

    hm	24. jan 2011	rev 1.1
    	improved performance
    *)

END_FUNCTION

(* ---- YEAR_OF_DATE.st ---- *)
FUNCTION YEAR_OF_DATE
    (*http://www.oscat.de/images/OSCATBasic/oscat_basic333_en.pdf#page=144*)
    YEAR_OF_DATE := UDINT_TO_INT((DATE_TO_UDINT(IDATE) + 43200) / 31557600 + 1970);

    (* revision history
    hm	4. aug 2006		rev 1.0
    	original version

    hm	1. okt 2007		rev 1.1
    	corrected error in algorithm
    	adjustment for S7 compatibility

    hm	23.12.2007		rev 1.2
    	changed code for better performance

    hm	7. apr. 2008	rev 1.3
    	deleted unused step7 code

    hm	7. oct. 2008	rev 1.4
    	renamed function (year) to YEAR_OF_DATE

    *)
END_FUNCTION

(* ---- _RMP_B.st ---- *)
FUNCTION_BLOCK _RMP_B
    (*http://www.oscat.de/images/OSCATBasic/oscat_basic333_en.pdf#page=255*)
    (* read system timer *)
    tx := UDINT_TO_TIME(T_PLC_MS());

    IF E AND init AND (DIR = last_dir) AND (BYTE_TO_USINT(RMP) <> SEL(DIR, 0, 255)) AND TR = tn THEN
    	RMP := FRMP_B(start, DIR, tx - tl, TR);
    ELSE
    	init := TRUE;
    	tl := tx;
    	tn := TR;
    	start := RMP;
    END_IF
    last_dir := DIR;

    (* revison history
    hm	22. oct. 2008	rev 1.0
    	original version

    hm	20. nov. 2008	rev 1.1
    	set default for E to be TRUE
    	added init

    hm	19. nov. 2011	rev 1.2
    	new code
    *)
END_FUNCTION_BLOCK

(* ---- _RMP_NEXT.st ---- *)
FUNCTION_BLOCK _RMP_NEXT
    (*http://www.oscat.de/images/OSCATBasic/oscat_basic333_en.pdf#page=255*)
    dirx(X := IN);

    t_lock(IN := FALSE, PT := TL);

    IF dirx.TU AND (OUT < IN) THEN
    	IF NOT xdir AND xen THEN t_lock(IN := TRUE); END_IF
    	xen := TRUE;
    	xdir := TRUE;
    ELSIF dirx.TD AND (OUT > IN) THEN
    	IF xdir AND xen THEN t_lock(IN := TRUE); END_IF
    	xen := TRUE;
    	xdir := FALSE;
    ELSIF xen THEN
    	IF (xdir AND (OUT >= IN)) OR (NOT xdir AND (OUT <= IN)) THEN
    		xen := FALSE;
    		IF TL > t#0s THEN t_lock(IN := TRUE); END_IF
    	END_IF
    END_IF

    IF NOT t_lock.Q AND xen THEN
    		UP := xdir;
    		DIR := xdir;
    		DN := NOT xdir;
    ELSE
    	UP := FALSE;
    	DN := FALSE;
    END_IF

    rmx(RMP := OUT, E := E AND (UP OR DN) , DIR := DIR, TR := SEL(DIR, TF, TR));

    (* revison history
    hm	23. nov. 2008	rev 1.0
    	original version

    hm	24. jan. 2009	rev 1.1
    	deleted unused vars tmp1, tmp2

    hm	20. feb. 2009	rev 1.2
    	improved algorithm
    	added TL

    hm	9. mar. 2009	rev 1.3
    	input E was ignored
    	removed double assignments

    hm	18. jul. 2009	rev 1.4
    	improved performance

    *)
END_FUNCTION_BLOCK

(* ---- _RMP_W.st ---- *)
FUNCTION_BLOCK _RMP_W
    (*http://www.oscat.de/images/OSCATBasic/oscat_basic333_en.pdf#page=256*)
    tx := T_PLC_MS();
    IF E AND init THEN
    	(* we need to set tl = tx when direction changes *)
    	IF DIR XOR last_dir THEN
    	 tl := tx;
    	 last_dir := DIR;
    	END_IF
    	(* check_elapsed time and calculate only if necessary *)
    	IF TR > t#0s THEN
    		step := UDINT_TO_DINT(SHL(tx-tl, 16) / TIME_TO_UDINT(TR));
    	ELSE
    		step := 65535;
    	END_IF
    	IF step > 0 THEN
    		(* perform the step on the ramp *)
    		tl := tx;
    		(* calculate the step response *)
    		IF NOT DIR THEN step := - step; END_IF
    		RMP := DINT_TO_WORD(LIMIT(0, WORD_TO_DINT(RMP) + step, 65535));
    	END_IF
    ELSE
    	tl := tx;
    	init := TRUE;
    END_IF

    (* revison history
    hm	22. oct. 2008	rev 1.0
    	original version

    hm	20. nov. 2008	rev 1.1
    	set default for E to be TRUE
    	added init

    *)
END_FUNCTION_BLOCK

(* ---- A_TRIG.st ---- *)
FUNCTION_BLOCK A_TRIG
    (*http://www.oscat.de/images/OSCATBasic/oscat_basic333_en.pdf#page=188*)
    D := IN - last_in;
    Q := ABS(D) > RES;
    IF Q THEN last_in := IN; END_IF
    D := IN - last_in;

    (* revision history

    hm 	16. jul. 2008	rev 1.0
    	original version released

    hm	25. oct. 2008	rev 1.1
    	code optimization
    	a_trig now also works for RES = 0

    *)
END_FUNCTION_BLOCK

(* ---- AIN1.st ---- *)
FUNCTION_BLOCK AIN1
    (*http://www.oscat.de/images/OSCATBasic/oscat_basic333_en.pdf#page=270*)
    (*Convert all dwords to udint as its not possible to do dword math*)
    _CODE_MIN := DWORD_TO_UDINT(CODE_MIN);
    _CODE_MAX := DWORD_TO_UDINT(CODE_MAX);
    (* extract ERROR bit *)
    ERROR := ((SHR(IN,ERROR_BIT) AND 16#0000_0001) = 1) OR (ERROR_CODE_EN AND ERROR_CODE = IN);
    IF ERROR THEN
    	OUT := ERROR_OUTPUT;
    	RETURN;
    END_IF

    (* strip off the data input *)
    tB := SHR(SHL(DWORD_TO_UDINT(IN), 31 - BIT_N), 31 - BIT_N + BIT_0);

    (* extract OVERFLOW bit *)
    OVERFLOW := ((SHR(IN,OVERFLOW_BIT) AND 16#0000_0001) = 1) OR (OVERFLOW_CODE_EN AND OVERFLOW_CODE = IN) OR (tB < _CODE_MIN OR tB > _CODE_MAX);
    IF OVERFLOW THEN
    	OUT := OVERFLOW_OUTPUT;
    	RETURN;
    END_IF

    (* extract SIGN bit *)
    SIGN := (SHR(IN,SIGN_BIT) AND 16#0000_0001) = 1;

    (* convert IN to OUT *)
    OUT := (UDINT_TO_REAL(tB - _CODE_MIN) * (OUT_MAX - OUT_MIN) / UDINT_TO_REAL(_CODE_MAX - _CODE_MIN) + OUT_MIN);
    IF SIGN THEN OUT := OUT * -1.0; END_IF

    (* revision history
    hm	23. feb 2008	rev 1.0
    	original version

    hm	16. mar 2008	rev 1.1
    	added type conversions to avoid warnngs under codesys 30

    hm	22. apr. 2008	rev 1.2
    	corrected ERROR IN formula when CODE_MIN was set
    	corrected ERROR when SIGN bit was used
    	optimized code for better performance

    hm	10. mar. 2009	rev 1.3
    	real constants updated to new systax using dot

    *)
END_FUNCTION_BLOCK

(* ---- ALARM_2.st ---- *)
FUNCTION_BLOCK ALARM_2
    (*http://www.oscat.de/images/OSCATBasic/oscat_basic333_en.pdf#page=333*)
    tmp := X - HYS * 0.5;
    IF tmp > LO_1 THEN Q1_LO := FALSE; END_IF
    IF tmp > LO_2 THEN Q2_LO := FALSE; END_IF
    IF tmp > HI_1 THEN Q1_HI := TRUE; END_IF
    IF tmp > HI_2 THEN Q2_HI := TRUE; END_IF
    tmp := tmp + HYS;
    IF tmp < LO_1 THEN Q1_LO := TRUE; END_IF
    IF tmp < LO_2 THEN Q2_LO := TRUE; END_IF
    IF tmp < HI_1 THEN Q1_HI := FALSE; END_IF
    IF tmp < HI_2 THEN Q2_HI := FALSE; END_IF

    (* revision history
    hm	19. may. 2008		rev 1.0
    	original version

    hm	11. mar. 2009	rev 1.1
    	improved code
    *)

END_FUNCTION_BLOCK

(* ---- ASTRO.st ---- *)
FUNCTION_BLOCK ASTRO
    (*http://www.oscat.de/images/OSCATBasic/oscat_basic333_en.pdf#page=354*)
    YAE :=	AE
    		+ M * 6.6845871535E-012
    		+ PC * 206265.0
    		+ LJ * 63240.0;
    YM := YAE * 149.597870E9;
    YPC := YAE * 4.8481322570E-006;
    YLJ := YAE * 1.5812776724E-005;

    (*
    Länge Meter M SI-Basiseinheit
    Astronomische Einheit* AE 1 AE = 149,597 870 · E9 M
    Parsec PC 1 PC = 206265 AE = 30,857 · E15 M
    Lichtjahr LJ 1 LJ = 9,460 530 · E15 M = 63240 AE = 0,306 59 PC
    Ångström Å 1 Å = E–l0 M
    typograph. Punkt p 1 p = 0,376 065 mm • im Druckereigewerbe
    inch** in 1 in = 2,54 · E–2 M = 25,4 mm***
    foot ft 1 ft = 0,3048 M = 30,48 cm
    yard yd 1 yd = 0,9144 M
    mile mile 1 mile = 1609,344 M
    Internat. Seemeile sm 1 sm = 1852 M
    Fathom fm 1 fm = 1,829 M • in der Seeschifffahrt
    *)

    (* revision history

    hm	27. mar. 2007	rev 1.0
    	original version

    hm	11. mar. 2009	rev 1.1
    	improved code

    *)

END_FUNCTION_BLOCK

(* ---- B_TRIG.st ---- *)
FUNCTION_BLOCK B_TRIG
    (*http://www.oscat.de/images/OSCATBasic/oscat_basic333_en.pdf#page=188*)
    Q := CLK XOR edge_;
    edge_ := CLK;

    (* revision history
    hm		4. aug. 2006	rev 1.0
    	original version

    *)
END_FUNCTION_BLOCK

(* ---- BAR_GRAPH.st ---- *)
FUNCTION_BLOCK BAR_GRAPH
    (*http://www.oscat.de/images/OSCATBasic/oscat_basic333_en.pdf#page=333*)
    IF NOT init THEN
    	init := TRUE;
    	IF LOG_SCALE THEN
    		temp := EXP(LN(TRIGGER_HIGH / TRIGGER_LOW) * 0.166666666666666666666);
    		T1 := TRIGGER_LOW * temp;
    		T2 := T1 * temp;
    		T3 := T2 * temp;
    		T4 := T3 * temp;
    		T5 := T4 * temp;
    	ELSE
    		temp := (TRIGGER_HIGH - TRIGGER_LOW) * 0.142857142;
    		T1 := TRIGGER_LOW + temp;
    		T2 := T1 + temp;
    		T3 := T2 + temp;
    		T4 := T3 + temp;
    		T5 := T4 + temp;
    	END_IF
    END_IF

    (* clear outputs before checking *)
    Q1 := FALSE;
    Q2 := FALSE;
    Q3 := FALSE;
    Q4 := FALSE;
    Q5 := FALSE;
    Q6 := FALSE;
    STATUS := 110;

    (* LOW, HIGH and ALARM can only be cleared with RST depending on ALARM_LOW and ALARM_HIGH *)
    IF NOT ALARM_LOW THEN LOW := FALSE; END_IF
    IF NOT ALARM_HIGH THEN HIGH := FALSE; END_IF
    IF RST THEN
    	ALARM := FALSE;
    	LOW := FALSE;
    	HIGH := FALSE;
    END_IF

    (* check and set outputs *)
    IF X < TRIGGER_LOW THEN
    	LOW := TRUE;
    	STATUS := 111;
    	IF ALARM_LOW THEN
    		ALARM := TRUE;
    		STATUS := 1;
    	END_IF
    ELSIF X < T1 THEN
    	Q1 := TRUE;
    ELSIF X < T2 THEN
    	Q2 := TRUE;
    ELSIF X < T3 THEN
    	Q3 := TRUE;
    ELSIF X < T4 THEN
    	Q4 := TRUE;
    ELSIF X < T5 THEN
    	Q5 := TRUE;
    ELSIF X < TRIGGER_HIGH THEN
    	Q6 := TRUE;
    ELSE
    	HIGH := TRUE;
    	STATUS := 112;
    	IF ALARM_HIGH THEN
    		ALARM := TRUE;
    		STATUS := 2;
    	END_IF
    END_IF

    (* revision history
    hm	22. feb 2007	rev 1.0
    	original version

    hm	2. dec 2007		rev 1.1
    	chaged code for better performance

    hm	6. jan 2008		rev 1.2
    	further performance improvement

    *)
END_FUNCTION_BLOCK

(* ---- BYTE_TO_BITS.st ---- *)
FUNCTION_BLOCK BYTE_TO_BITS
    (*http://www.oscat.de/images/OSCATBasic/oscat_basic333_en.pdf#page=216*)
    B0 := IN.0;
    B1 := IN.1;
    B2 := IN.2;
    B3 := IN.3;
    B4 := IN.4;
    B5 := IN.5;
    B6 := IN.6;
    B7 := IN.7;

    (* revision history
    hm		4. aug 2006	rev 1.0
    	original version

    hm		16. mar 2008	rev 1.1
    	renamed from byte_to_bit to byte_to_bits for compatibility reasons

    *)
END_FUNCTION_BLOCK

(* ---- CALENDAR_CALC.st ---- *)
FUNCTION_BLOCK CALENDAR_CALC
    (*http://www.oscat.de/images/OSCATBasic/oscat_basic333_en.pdf#page=114*)
    IF XCAL.UTC <> last THEN
    	(* run once per second *)
    	(* update utc last calculated  *)
    	last := XCAL.UTC;
    	utod := DT_TO_TOD(XCAL.UTC);

    	(* calculate ltc from utc *)
    	XCAL.LOCAL_DT := UTC_TO_LTIME(XCAL.UTC, XCAL.DST_EN, XCAL.OFFSET);
    	XCAL.LOCAL_DATE := DT_TO_DATE(XCAL.LOCAL_DT);
    	XCAL.LOCAL_TOD := DT_TO_TOD(XCAL.LOCAL_DT);
    	dtemp := DAY_OF_DATE(XCAL.LOCAL_DATE);
    	XCAL.NIGHT := XCAL.LOCAL_TOD < XCAL.SUN_RISE OR XCAL.LOCAL_TOD > XCAL.SUN_SET;

    	(* run once per hour *)
    	tmp := HOUR(XCAL.LOCAL_TOD);
    	IF  tmp <> last_hour THEN
    		XCAL.DST_ON := DST(XCAL.UTC) AND XCAL.DST_EN;
    		last_hour := tmp;
    	END_IF

    	(* run once per day *)
    	IF dtemp <> last_day THEN
    		last_day := dtemp;
    		(* a new day has started, recalculate daily events *)
    		XCAL.YEAR := YEAR_OF_DATE(XCAL.LOCAL_DATE);
    		XCAL.MONTH := MONTH_OF_DATE(XCAL.LOCAL_DATE);
    		XCAL.DAY := DAY_OF_MONTH(XCAL.LOCAL_DATE);
    		XCAL.WEEKDAY := DAY_OF_WEEK(XCAL.LOCAL_DATE);
    		holy(DATE_IN := XCAL.LOCAL_DATE, LANGU := XCAL.LANGUAGE, HOLIDAYS := HOLIDAYS);
    		XCAL.HOLIDAY := holy.Y;
    		XCAL.HOLY_NAME := holy.NAME;
    		sun(LATITUDE := XCAL.LATITUDE, LONGITUDE := XCAL.LONGITUDE, UTC := DT_TO_DATE(XCAL.UTC), H := H);
    		XCAL.SUN_RISE := DINT_TO_TOD(TOD_TO_DINT(sun.SUN_RISE) + XCAL.OFFSET * 60000 + SEL(XCAL.DST_ON,DINT#0,3600000));
    		XCAL.SUN_SET := DINT_TO_TOD(TOD_TO_DINT(sun.SUN_SET) + XCAL.OFFSET * 60000 + SEL(XCAL.DST_ON,DINT#0,3600000));
    		XCAL.SUN_MIDDAY := DINT_TO_TOD(TOD_TO_DINT(sun.MIDDAY) + XCAL.OFFSET * 60000 + SEL(XCAL.DST_ON,DINT#0,3600000));
    		XCAL.SUN_HEIGTH := sun.SUN_DECLINATION;
    		XCAL.WORK_WEEK := WORK_WEEK(XCAL.LOCAL_DATE);
    	END_IF

    	(* calculate the suns position every 10 seconds when SPE = TRUE *)
    	IF SPE AND XCAL.UTC -  plast >= t#25s THEN
    		plast := last;
    		pos(LATITUDE := XCAL.LATITUDE, LONGITUDE := XCAL.LONGITUDE, UTC := XCAL.UTC);
    		XCAL.SUN_HOR := pos.B;
    		XCAL.SUN_VER := pos.HR;
    	END_IF
    END_IF

    (* revision history

    hm 23. oct. 2008	rev 1.0
    	original version

    hm	8. feb. 2009	rev 1.1
    	night was calculated wrong
    	added sun position data

    hm	10. mar. 2009	rev 1.2
    	added work_week, sun_midday, sun_heigth
    	sun_position will only be calculated evey 25 seconds
    	dst will only become true when dst_en = true

    hm	23. jan 2010	rev 1.3
    	sun_rise, sun_set and sun_midday are now calculated in local time

    hm	18. jan. 2011	rev 1.4
    	added input HOLIDAYS to specify local HOLIDAYS
    	changed call for function sun_time

    hm	2. feb. 2011	rev 1.5
    	added input H to specify twilight

    hm	6. apr. 2011	rev 1.6
    	night was calculated wrong

    HM 3. Feb 2021    rev 1.7
       chaged LDT >> LOCAL_DT, LDATE >> LOCAL_DT, LTOD >> LOCAL_TOD

    *)
END_FUNCTION_BLOCK

(* ---- CALIBRATE.st ---- *)
FUNCTION_BLOCK CALIBRATE
    (*http://www.oscat.de/images/OSCATBasic/oscat_basic333_en.pdf#page=337*)
    (* check for calibration *)
    IF CO THEN
    	offset := Y_OFFSET - X;
    ELSIF CS THEN
    	Scale := Y_SCALE / (X + offset);
    END_IF
    (* calculate output *)
    Y := (X + offset) * Scale;

    (* revision history
    hm 22.2.2007		rev 1.2
    	changed VAR RETAIN PERSISTENT to VAR RETAIN for better compatibility
    	wago lon contollers do not support persisitent

    hm	11. mar. 2009	rev 1.3
    	changed real constants to use dot syntax

    *)
END_FUNCTION_BLOCK

(* ---- CLICK_CNT.st ---- *)
FUNCTION_BLOCK CLICK_CNT
    (*http://www.oscat.de/images/OSCATBasic/oscat_basic333_en.pdf#page=189*)
    (* Q shall only be active for one cycle only *)
    Q := FALSE;

    IF IN AND NOT edge_ AND NOT tx.Q THEN
    	(* a rising edge_ on IN sets the counter to 0 *)
    	cnt := 0;
    ELSIF tx.Q AND NOT IN AND edge_ THEN
    	(* count falling edges when tp.Q is true *)
    	cnt := cnt + 1;
    ELSIF NOT tx.Q THEN
    	Q := cnt = N;
    	cnt := -1;
    END_IF

    (* remember the status of IN *)
    edge_ := IN;
    tx(IN := IN, PT := TC);

    (* revision history

    hm 	16. jul. 2008	rev 1.0
    	original version released

    *)
END_FUNCTION_BLOCK

(* ---- CLICK_DEC.st ---- *)
FUNCTION_BLOCK CLICK_DEC
    (*http://www.oscat.de/images/OSCATBasic/oscat_basic333_en.pdf#page=190*)
    (* Q shall only be active for one cycle only *)
    IF IN = FALSE THEN
    	Q0 := FALSE;
    	Q1 := FALSE;
    	Q2:= FALSE;
    	Q3 := FALSE;
    END_IF

    IF IN AND NOT edge_ AND NOT tx.Q THEN
    	(* a rising edge_ on IN sets the counter to 0 *)
    	cnt := 0;
    ELSIF tx.Q AND NOT IN AND edge_ THEN
    	(* count falling edges when tp.q is true *)
    	cnt := cnt + 1;
    ELSIF NOT tx.Q THEN
    	CASE cnt OF
    		0 : Q0 := TRUE;
    		1 : Q1 := TRUE;
    		2 : Q2 := TRUE;
    		3 : Q3 := TRUE;
    	END_CASE
    	cnt := -1;
    END_IF

    (* remember the status of IN *)
    edge_ := IN;
    tx(IN := IN, PT := TC);

    (* revision history

    hm 17. jul. 2008	rev 1.0
    	original version released

    hm	14. mar. 2009	rev 1.1
    	removed double assignments

    *)
END_FUNCTION_BLOCK

(* ---- CLK_DIV.st ---- *)
FUNCTION_BLOCK CLK_DIV
    (*http://www.oscat.de/images/OSCATBasic/oscat_basic333_en.pdf#page=190*)
    IF RST THEN
    	cnt:= 0;
    	Q0 := 0;
    	Q1 := 0;
    	Q2 := 0;
    	Q3 := 0;
    	Q4 := 0;
    	Q5 := 0;
    	Q6 := 0;
    	Q7 := 0;
    ELSIF CLK THEN
    	cnt:= cnt +1;
    	Q0 := cnt.0;
    	Q1 := cnt.1;
    	Q2 := cnt.2;
    	Q3 := cnt.3;
    	Q4 := cnt.4;
    	Q5 := cnt.5;
    	Q6 := cnt.6;
    	Q7 := cnt.7;
    END_IF

    (* revision history
    hm	4. aug. 2006	rev 1.0
    	original version

    hm	2. jan 2008		rev 1.1
    	improved performance

    *)
END_FUNCTION_BLOCK

(* ---- CLK_N.st ---- *)
FUNCTION_BLOCK CLK_N
    (*http://www.oscat.de/images/OSCATBasic/oscat_basic333_en.pdf#page=192*)
    stime := SHR(T_PLC_MS(),N);
    clk := stime.0;
    Q := clk XOR edge_;
    edge_ := clk;

    (* revision history
    hm	16. dec 2007		rev 1.0
    	original version

    *)
END_FUNCTION_BLOCK

(* ---- CLK_PRG.st ---- *)
FUNCTION_BLOCK CLK_PRG
    (*http://www.oscat.de/images/OSCATBasic/oscat_basic333_en.pdf#page=192*)
    (* read system time *)
    tx := UDINT_TO_TIME(T_PLC_MS());

    (* initialize on startup *)
    IF NOT init THEN
    	init := TRUE;
    	last := tx - PT;
    END_IF

    (* generate output pulse when next_pulse is reached *)
    Q := tx - last >= PT;
    IF Q THEN last := tx; END_IF

    (* revision hiostory

    hm 25 feb 2007	rev 1.1
    	rewritten code for higher performance
    	PT can now be changed during runtime

    hm	17. sep 2007	rev 1.2
    	replaced time() with t_plc_ms() for compatibility reasons

    hm	25. oct. 2008	rev 1.3
    	optimized code

    *)
END_FUNCTION_BLOCK

(* ---- CLK_PULSE.st ---- *)
FUNCTION_BLOCK CLK_PULSE
    (*http://www.oscat.de/images/OSCATBasic/oscat_basic333_en.pdf#page=193*)
    tx := T_PLC_MS();		(* read system *)
    Q := FALSE;				(* reset Q we generate pulses only for one cycle *)
    RUN := CNT < N;

    IF NOT init OR RST THEN
    	init := TRUE;
    	CNT := 0;
    	tn := tx - TIME_TO_UDINT(PT);
    	RUN := FALSE;
    ELSIF (CNT < N OR N = 0) AND tx - tn >= TIME_TO_UDINT(PT) THEN		(* generate a pulse *)
    	CNT := CNT + 1;
    	Q := TRUE;
    	tn := tn + TIME_TO_UDINT(PT);
    END_IF

    (* revision history
    hm		4. aug 2006		rev 1.0
    	original version

    hm		17. sep 2007	rev 1.1
    	replaced time() with T_PLC_S() for compatblity reasons

    hm		16. feb. 2011	rev 1.2
    	fixed an error when timer overflows
    *)
END_FUNCTION_BLOCK

(* ---- CONTROL_SET1.st ---- *)
FUNCTION_BLOCK CONTROL_SET1
    (*http://www.oscat.de/images/OSCATBasic/oscat_basic333_en.pdf#page=377*)
    IF PI AND PID THEN
    	KP := 0.0;
    	TN := 0.0;
    	TV := 0.0;
    ELSIF PID THEN
    	KP := PID_K * KT;
    	TN := PID_TN * TT;
    	TV := PID_TV * TT;
    ELSIF PI THEN
    	KP := PI_K * KT;
    	TN := PI_TN * TT;
    ELSE
    	KP := P_K * KT;
    END_IF

    (* KI and KD are calculated *)
    IF TN > 0.0 THEN KI := KP / TN; ELSE KI := 0.0; END_IF
    KD := KP * TV;

    (* revision history
    hm	4. nov 2007	rev 1.0
    	original version

    hm	11. mar. 2009	rev 1.1
    	real constants updated to new systax using dot

    *)
END_FUNCTION_BLOCK

(* ---- CONTROL_SET2.st ---- *)
FUNCTION_BLOCK CONTROL_SET2
    (*http://www.oscat.de/images/OSCATBasic/oscat_basic333_en.pdf#page=379*)
    IF TU > 0.0 AND KS > 0.0 THEN TX := TG / TU / KS; END_IF
    IF PI AND PID THEN
    	KP := 0.0;
    	TN := 0.0;
    	TV := 0.0;
    ELSIF PID THEN
    	KP := PID_K * TX;
    	TN := PID_TN * TU;
    	TV := PID_TV * TU;
    ELSIF PI THEN
    	KP := PI_K * TX;
    	TN := PI_TN * TU;
    ELSE
    	KP := P_K * TX;
    END_IF

    (* KI and KD are calculated *)
    IF TN > 0.0 THEN KI := KP / TN; ELSE KI := 0.0; END_IF
    KD := KP * TV;

    (* revision history
    hm	4. nov 2007	rev 1.0
    	original version

    hm	11. mar. 2009	rev 1.1
    	real constants updated to new systax using dot

    *)
END_FUNCTION_BLOCK

(* ---- COUNT_BR.st ---- *)
FUNCTION_BLOCK COUNT_BR
    (*http://www.oscat.de/images/OSCATBasic/oscat_basic333_en.pdf#page=236*)
    IF RST THEN
    	CNT := 0;
    ELSIF SET THEN
    	CNT := LIMIT(0,IN,MX);
    ELSIF UP AND NOT last_up THEN
    	CNT := INT_TO_BYTE(INC(BYTE_TO_USINT(CNT),BYTE_TO_USINT(STEP),BYTE_TO_USINT(MX)));
    ELSIF DN AND NOT last_dn THEN
    	CNT := INT_TO_BYTE(INC(BYTE_TO_USINT(CNT),-BYTE_TO_USINT(STEP),BYTE_TO_USINT(MX)));
    END_IF
    last_up := UP;
    last_dn := DN;

    (* revision history
    hm	16. jan 2008	rev 1.0
    	original version

    *)
END_FUNCTION_BLOCK

(* ---- COUNT_DR.st ---- *)
FUNCTION_BLOCK COUNT_DR
    (*http://www.oscat.de/images/OSCATBasic/oscat_basic333_en.pdf#page=237*)
    _MX := DWORD_TO_UDINT(MX);
    _STEP := DWORD_TO_UDINT(STEP);
    _IN := DWORD_TO_UDINT(IN);
    IF RST THEN
    	_CNT := 0;
    ELSIF SET THEN
    	_CNT := LIMIT(0,_IN,_MX);
    ELSIF UP AND NOT last_up THEN
    	IF _STEP > _MX - _CNT THEN
    		_CNT := _CNT - _MX + _STEP - 1;
    	ELSE
    		_CNT := _CNT + _STEP;
    	END_IF
    ELSIF DN AND NOT last_dn THEN
    	IF _STEP > _CNT THEN
    		_CNT := _CNT - _STEP + _MX + 1;
    	ELSE
    		_CNT := _CNT - _STEP;
    	END_IF
    END_IF
    last_up := UP;
    last_dn := DN;
    CNT := UDINT_TO_DWORD(_CNT);
    (* revision history
    hm	12. jun 2008	rev 1.0
    	original version

    hm	20. jan. 2011	rev 1.1
    	corrected init value of MX to 16#FFFFFFFF

    *)
END_FUNCTION_BLOCK

(* ---- CTRL_OUT.st ---- *)
FUNCTION_BLOCK CTRL_OUT
    (*http://www.oscat.de/images/OSCATBasic/oscat_basic333_en.pdf#page=381*)
    Y := SEL(MANUAL, CI, MAN_IN) + OFFSET;

    (* Limit the output *)
    IF Y > LIM_L AND Y < LIM_H THEN
    	LIM := FALSE;
    ELSE
    	Y := LIMIT(LIM_L, Y, LIM_H);
    	LIM := TRUE;
    END_IF

    (* revision history
    hm 	2. jun. 2008 	rev 1.0
    	original version

    hm	5. nov. 2008	rev 1.1
    	optimized code
    *)
END_FUNCTION_BLOCK

(* ---- CTRL_PI.st ---- *)
FUNCTION_BLOCK CTRL_PI
    (*http://www.oscat.de/images/OSCATBasic/oscat_basic333_en.pdf#page=382*)
    DIFF := CTRL_IN(SET, ACT, SUP);
    pi(IN := DIFF, KP := KP, KI := KI, LIM_L := LL, LIM_H := LH, RST := RST);
    co(CI := pi.Y, OFFSET := OFS, MAN_IN := M_I, LIM_L := LL, LIM_H := LH, MANUAL := MAN);
    Y := co.Y;
    LIM := co.LIM;

    (* revision history
    hm 	31.10.2007 		rev 1.0
    	original version

    hm	3.11.2007		rev 1.1
    	added noise input to filter noise
    	added output DIFF
    	SET limit output false when output is within limits
    	overfolw was not SET correctly

    hm	5. jan 2008		rev 1.2
    	improved performance

    hm	20. jun. 2008	rev 2.0
    	rewritten using new modular approach

    *)
END_FUNCTION_BLOCK

(* ---- CTRL_PID.st ---- *)
FUNCTION_BLOCK CTRL_PID
    (*http://www.oscat.de/images/OSCATBasic/oscat_basic333_en.pdf#page=384*)
    DIFF := CTRL_IN(SET, ACT, SUP);
    pid(IN := DIFF, KP := KP, TN := TN, TV := TV, LIM_L := LL, LIM_H := LH, RST := RST);
    co(CI := pid.Y, OFFSET := OFS, MAN_IN := M_I, LIM_L := LL, LIM_H := LH, MANUAL := MAN);
    Y := co.Y;
    LIM := co.LIM;

    (* revision history

    hm 1.12.2006	 	rev 1.1
    	changed algorithm to trapezregel for higher accuracy.

    hm 3.1.2007		rev 1.2
    	added integ_band to select when the integrator is active.

    hm	3.3.2007		rev 1.3
    	added default values to inputs KP, TN, TV, LIMIT_L und LIMIT_H.

    hm 31.oct 2007	rev 1.4
    	total rewrite of the module to avoid failures when one of the limits is 0

    hm	3.11.2007	rev 1.5
    	added noise input to filter noise
    	added output DIFF
    	SET limit output false when output is within limits
    	overfolw was not SET correctly

    hm	5. jan 2008	rev 1.6
    	improved code for better performance
    *)
END_FUNCTION_BLOCK

(* ---- CTRL_PWM.st ---- *)
FUNCTION_BLOCK CTRL_PWM
    (*http://www.oscat.de/images/OSCATBasic/oscat_basic333_en.pdf#page=386*)
    PW(F := F, DC := SEL(MANUAL,CI,MAN_IN));
    Q := PW.Q;

    (* revision history
    hm 3. jun. 2008 	rev 1.0
    	original version

    hm	21. oct. 2008	rev 1.1
    	optimized code

    *)
END_FUNCTION_BLOCK

(* ---- CYCLE_4.st ---- *)
FUNCTION_BLOCK CYCLE_4
    (*http://www.oscat.de/images/OSCATBasic/oscat_basic333_en.pdf#page=194*)
    (* read system timer *)
    tx := UDINT_TO_TIME(T_PLC_MS());
    (* init on first cycle *)
    IF NOT init THEN
    	init := TRUE;
    	last := tx;
    END_IF

    IF E THEN
    	IF SL THEN
    		(* when SX > 0 then the STATE SX is forced to start *)
    		STATE:= LIMIT(0,SX,3);
    		last := tx;
    		(* this is to avoid to reset SX from the calling programm it does work fine on codesys but i am not sure about other systems, because we are writing to an input *)
    		SL := FALSE;
    	ELSE
    		CASE STATE OF
    			0 :	(* wait for T0 and switch to next cycle *)
    				IF tx - last >= T0 THEN
    					STATE := 1;
    					last := tx;
    				END_IF
    			1 : (* wait for T1 over 1st cycle *)
    				IF tx - last >= T1 THEN
    					STATE := 2;
    					last := tx;
    				END_IF
    			2 : (* wait for T1 over 1st cycle *)
    				IF tx - last >= T2 THEN
    					STATE := 3;
    					last := tx;
    				END_IF
    			3 : (* wait for T2 over 2nd cycle *)
    				IF tx - last >= T3 THEN
    					IF S0 THEN STATE := 0; END_IF (* if S0 is false, the sequence stops at STATE 3 *)
    					last := tx;
    				END_IF
    		END_CASE
    	END_IF
    ELSE
    	STATE := 0;
    	last := tx;
    END_IF

    (*
    hm	3. nov. 2008	rev 1.0
    	original version

    *)
END_FUNCTION_BLOCK

(* ---- CYCLE_TIME.st ---- *)
FUNCTION_BLOCK CYCLE_TIME
    (*http://www.oscat.de/images/OSCATBasic/oscat_basic333_en.pdf#page=338*)
    tx := UDINT_TO_TIME(T_PLC_MS()) - last_cycle;
    IF RST THEN
    	CT_MIN := t#10h;
    	CT_MAX := t#0ms;
    	CYCLES := 0;
    ELSIF last_cycle > t#0s THEN
    	IF tx < CT_MIN THEN CT_MIN := tx;
    	ELSIF tx > CT_MAX THEN CT_MAX := tx;
    	END_IF
    	CT_LAST := tx;
    ELSIF CT_MIN = t#0s THEN
    	CT_MIN := t#0s - t#1ms;
    END_IF
    IF init THEN
    	SYSTIME := SYSTIME + tx;
    		IF SYSTIME >= t#1d THEN
    			SYSTIME := SYSTIME - t#1d;
    			SYSDAYS := SYSDAYS + 1;
    		END_IF
    END_IF
    init := TRUE;
    last_cycle := last_cycle + tx;
    CYCLES := CYCLES + 1;

    (*	revision history
    hm 12.12.2006		rev 1.1
    	added CYCLES output, a UDINT cycle counter.
    hm 10.3.2007			rev 1.2
    	changed initialization of CT_MIN to t#10h for compatibility with siemens s7

    hm	16.9.2007		rev 1.2
    	changed Time() in T_PLC_MS() for compatibility resons

    *)
END_FUNCTION_BLOCK

(* ---- D_TRIG.st ---- *)
FUNCTION_BLOCK D_TRIG
    (*http://www.oscat.de/images/OSCATBasic/oscat_basic333_en.pdf#page=195*)
    Q := IN <> last_in;
    X := UDINT_TO_DWORD(DWORD_TO_UDINT(IN) - DWORD_TO_UDINT(last_in));
    last_in := IN;

    (* revision history

    hm 	4.09.2007		rev 1.0
    	original version released

    hm	19. feb. 2008	rev 1.1
    	performance improvement
    *)
END_FUNCTION_BLOCK

(* ---- DCF77.st ---- *)
FUNCTION_BLOCK DCF77
    (*http://www.oscat.de/images/OSCATBasic/oscat_basic333_en.pdf#page=119*)
    (* if TP was SET it should only be active for 1 cycle *)
    TP := FALSE;

    (* read system time *)
    t1 := UDINT_TO_TIME(T_PLC_MS());
    tx := t1 - last;

    IF REC XOR edge_ THEN
    	edge_ := REC;
    	IF NOT REC AND tx > t#1700ms AND tx < t#2000ms THEN
    		(* start condition reached *)
    		state := 0;
    		TP := NOT ERROR;
    	ELSIF NOT REC AND tx > t#700ms AND tx < t#1000ms THEN
    		(* second switch detected *)
    		IF state < 58 THEN state := state +1; ELSE state := 0; END_IF
    	ELSIF REC AND tx  < t#120ms THEN
    		(* bit 0 detected  *)
    		bits[state] := 0;
    	ELSIF REC AND tx > t#120ms AND tx < t#250ms THEN
    		(* bit 1 detected *)
    		bits[state] := 1;
    	ELSE
    		(* ERROR condition received signal is not valid *)
    		ERROR := TRUE;
    		state := 0;
    	END_IF
    	last := last + tx;
    	IF REC AND state = 58 THEN
    		ERROR := FALSE;

    		(* decode the bits and check for possible errors *)
    		IF bits[0] OR NOT (bits[17] XOR bits[18]) OR NOT bits[20] THEN ERROR := TRUE; END_IF
    		(* decode minute *)
    		minute := 0;
    		minute.0 := bits[21];
    		minute.1 := bits[22];
    		minute.2 := bits[23];
    		minute.3 := bits[24];
    		IF bits[25] THEN minute := minute + 10; END_IF
    		IF bits[26] THEN minute := minute + 20; END_IF
    		IF bits[27] THEN minute := minute + 40; END_IF
    		IF minute > 59 OR (bits[21] XOR bits[22] XOR bits[23] XOR bits[24] XOR bits[25] XOR bits[26] XOR bits[27] XOR bits[28]) THEN ERROR := TRUE; END_IF

    		(* decode hour *)
    		hour := 0;
    		hour.0 := bits[29];
    		hour.1 := bits[30];
    		hour.2 := bits[31];
    		hour.3 := bits[32];
    		IF bits[33] THEN hour := hour + 10; END_IF
    		IF bits[34] THEN hour := hour +20; END_IF
    		IF hour > 23 OR (bits[29] XOR bits[30] XOR bits[31] XOR bits[32] XOR bits[33] XOR bits[34] XOR bits[35]) THEN ERROR := TRUE; END_IF

    		(* decode day of month *)
    		day := 0;
    		day.0 := bits[36];
    		day.1 := bits[37];
    		day.2 := bits[38];
    		day.3 := bits[39];
    		IF bits[40] THEN day := day + 10; END_IF
    		IF bits[41] THEN day := day + 20; END_IF
    		IF day > 31 THEN ERROR := TRUE; END_IF

    		(* decode day of week *)
    		WDAY := 0;
    		WDAY.0 := bits[42];
    		WDAY.1 := bits[43];
    		WDAY.2 := bits[44];
    		IF WDAY > 7 OR WDAY < 1 THEN ERROR := TRUE; END_IF

    		(* decode month *)
    		month := 0;
    		month.0 := bits[45];
    		month.1 := bits[46];
    		month.2 := bits[47];
    		month.3 := bits[48];
    		IF bits[49] THEN month := month +10; END_IF
    		IF month > 12 THEN ERROR := TRUE; END_IF

    		(* decode year *)
    		year := 0;
    		year.0 := bits[50];
    		year.1 := bits[51];
    		year.2 := bits[52];
    		year.3 := bits[53];
    		IF bits[54] THEN year := year + 10; END_IF
    		IF bits[55] THEN year := year + 20; END_IF
    		IF bits[56] THEN year := year + 40; END_IF
    		IF bits[57] THEN year := year + 80; END_IF

    		(* check parity for bits 36 to 58 *)
    		cnt := 0;
    		FOR i := 36 TO 58 DO IF bits[i] THEN cnt := cnt + 1; END_IF END_FOR
    		IF NOT EVEN(cnt) THEN ERROR := TRUE; END_IF

    		(* time must be valid for two cycles to clear ERROR flag *)
    		IF NOT ERROR THEN
    			(* SET outputs *)
    			old_time := mez;
    			IF year >= 70 THEN year := year + 1900; ELSE year := year + 2000; END_IF
    			mez := SET_DT(year,month,day,hour,minute,0);
    			DS := bits[17];
    			IF DS THEN
    				utc := UDINT_TO_DT(DT_TO_UDINT(mez) - 7200);
    			ELSE
    				utc := UDINT_TO_DT(DT_TO_UDINT(mez) - 3600);
    			END_IF

    			(* SET trigger signal only if the receiver has received 2 successive minutes *)
    			IF mez <> old_time + t#1m THEN ERROR := TRUE ; END_IF
    		END_IF
    	END_IF
    END_IF

    (* this portion implements a free running clock which is triggered by the dcf77 signal *)
    tz := UDINT_TO_TIME(INT_TO_UDINT(ABS(TIME_OFFSET))* 3600000);

    (* input SDT is copied to utc at first power up *)
    IF NOT init OR SET THEN
    	init := TRUE;
    	utc := SDT;
    	TP := TRUE;
    	DS := DSI;
    END_IF

    IF TP THEN
    	RTC := utc;
    	IF DS AND DST_EN THEN
    		IF TIME_OFFSET < 0 THEN	RTC1 := RTC - tz + t#1h; ELSE RTC1 := RTC + tz + t#1h; END_IF
    	ELSE
    		IF TIME_OFFSET < 0 THEN RTC1 := RTC - tz; ELSE RTC1 := RTC + tz; END_IF
    	END_IF
    	SYNC := TRUE;
    	last_sync := last;
    	ty := last;
    ELSIF RTC > UDINT_TO_DT(0) AND t1 - ty >= t#1s THEN
    	RTC := RTC + t#1s;
    	RTC1 := RTC1 + t#1s;
    	ty := ty + t#1s;
    	SYNC := ty - last_sync < SYNC_TIMEOUT AND last_sync > UDINT_TO_TIME(0);
    	WDAY := DAY_OF_WEEK(DT_TO_DATE(RTC1));
    	DS := DST_EN AND DST(utc);
    END_IF
    MSEC := TIME_TO_INT(t1 - ty);

    (* decode information
    bits		content
    0			Bitwert immer 0
    1 bis 14	reserviert für Betriebsinformationen (nicht für DCF77-Nutzer bestimmt)
    15			Rufbit für Alarmierung der PTB-Mitarbeiter
    			(bis Mai 2003: Bitwert = 0 falls normale Antenne in Verwendung; 1 = Backupantenne)
    16			Bitwert = 1 falls ein Wechsel von mez nach MESZ oder umgekehrt bevorsteht; Dauer der Anzeige: 1 Stunde
    17 + 18	gültige Zeit = mez, falls Bit 17=0 und Bit 18=1
    			gültige Zeit = MESZ, falls Bit 17=1 und Bit 18=0
    19			Bitwert = 1 falls innerhalb den nächsten 59 Minuten eine Schaltsekunde angeordnet ist. Beim Einfügen einer Schaltsekunde wird anstelle der 59. die 60. Sekundenmarke weggelassen und in der 58. erfolgt ausnahmsweise ein Trägerabfall.
    20			Startbit für Zeitinformation (immer 1)
    21 - 27		1, 2, 4, 8, 10, 20, 40 Minuten (bitweise Addition)
    28			Prüfbit (gerade Parität) für die bits 21-27
    29 - 34		1, 2, 4, 8, 10, 20 Stunden (bitweise Addition)
    35			Prüfbit (gerade Parität) für die bits 29-34
    36 - 41		Tagesnummer im aktuellen Monat: 1, 2, 4, 8, 10, 20 (bitweise Addition)
    42 - 44		Tagesnummer in der aktuellen Woche: 1, 2, 4 (bitweise Addition)
    45 - 49		Monatsnummer: 1, 2, 4, 8, 10 (bitweise Addition)
    50 - 57		Jahr (zweistellig): 1, 2, 4, 8, 10, 20, 40, 80 (bitweise Addition)
    58			Prüfbit (gerade Parität) füR die bits 36-57

    *)
    (* revision history

    hm 2.feb 2007		rev 1.1
    	change WDAY and dst outputs when there is no dcf reception

    hm	26.feb 2007		rev 1.2
    	changed statements where t#1h would be substracted from DT.
    	under certain conditions the compiler would crash translating this statement

    hm	17. sep 2007	rev 1.3
    	replaced time() with T_PLC_MS() for compatibility reasons

    hm	24. oct 2007		rev 1.4
    	changed dst calculation because function dst was upgraded no ERROR in DCF77 only a change in DST

    hm	12. nov 2007		rev 1.5
    	changed TIME_OFFSET from time to integer to allow for negative offset time zones

    hm	8. dec 2007		rev 1.6
    	corrected an ERROR in time_zone calculation

    hm 23. jan 2008		rev 1.7
    	added SDT input which is used to initialize RTC and RTC1 during first cycle.

    hm 16. mar 2008		rev 1.8
    	changed output weekday to WDAY and dst to DS for compatibility reasons

    hm	19. apr. 2008	rev 1.9
    	added input DSI to allow to SET daylight savings time when SDT is TRUE.
    	added asynchronous SET input

    hm	7. oct. 2008	rev 1.10
    	changed function weekday to day_of_week

    *)

END_FUNCTION_BLOCK

(* ---- DEAD_BAND_A.st ---- *)
FUNCTION_BLOCK DEAD_BAND_A
    (*http://www.oscat.de/images/OSCATBasic/oscat_basic333_en.pdf#page=393*)
    (* filter the input signal *)
    tp1(IN := X, T:= T);

    (* filter the HF portion to generate a stable L *)
    tp2(IN := ABS(tp1.OUT - X), T := MULTIME(T, 4.0));

    (* now we determine L which is half the width of the dead band *)
    L := MIN(KL * tp2.OUT, LM);

    IF X > L THEN
    	Y := X - L;
    ELSIF X < -L THEN
    	Y := X + L;
    ELSE
    	Y := 0.0;
    END_IF

    (* revision history
    hm	14. jun. 2008	rev 1.0
    	original version

    hm	11. mar. 2009	rev 1.1
    	real constants updated to new systax using dot

    *)
END_FUNCTION_BLOCK

(* ---- DEAD_ZONE2.st ---- *)
FUNCTION_BLOCK DEAD_ZONE2
    (*http://www.oscat.de/images/OSCATBasic/oscat_basic333_en.pdf#page=395*)
    IF ABS(X) > L THEN
    	Y := X;
    ELSIF Y > 0.0 THEN
    	Y := L;
    ELSE
    	Y := -L;
    END_IF

    (* revision history

    hm	12. feb. 2007	rev 1.0
    	original version

    hm	11. mar. 2009	rev 1.1
    	real constants updated to new systax using dot

    *)

END_FUNCTION_BLOCK

(* ---- DEC_2.st ---- *)
FUNCTION_BLOCK DEC_2
    (*http://www.oscat.de/images/OSCATBasic/oscat_basic333_en.pdf#page=222*)
    Q0 := D AND NOT A;
    Q1 := D AND A;

    (* revision history
    hm 3.3.2007	rev 1.1
    	rewritten in ST for better compatibility

    *)
END_FUNCTION_BLOCK

(* ---- DEC_4.st ---- *)
FUNCTION_BLOCK DEC_4
    (*http://www.oscat.de/images/OSCATBasic/oscat_basic333_en.pdf#page=222*)
    Q0 := D AND NOT A0 AND NOT A1;
    Q1 := D AND A0 AND NOT A1;
    Q2 := D AND NOT A0 AND A1;
    Q3 := D AND A0 AND A1;

    (* revision history
    hm 3.3.2007	rev 1.1
    	rewritten in ST for better compatibility

    *)
END_FUNCTION_BLOCK

(* ---- DEC_8.st ---- *)
FUNCTION_BLOCK DEC_8
    (*http://www.oscat.de/images/OSCATBasic/oscat_basic333_en.pdf#page=223*)
    X.0 := A0; X.1 := A1; X.2 := A2;

    Q0 := FALSE;
    Q1 := FALSE;
    Q2 := FALSE;
    Q3 := FALSE;
    Q4 := FALSE;
    Q5 := FALSE;
    Q6 := FALSE;
    Q7 := FALSE;

    CASE X OF
    	0 : Q0 := D;
    	1 : Q1 := D;
    	2 : Q2 := D;
    	3 : Q3 := D;
    	4 : Q4 := D;
    	5 : Q5 := D;
    	6 : Q6 := D;
    	7 : Q7 := D;
    END_CASE

    (* revision history
    hm 3. mar. 2007	rev 1.1
    	rewritten in ST for better compatibility

    hm	26. oct. 2008	rev 1.2
    	code optimized

    hm	28. mar. 2009	rev 1.3
    	replaced multiple assignments
    *)
END_FUNCTION_BLOCK

(* ---- DELAY.st ---- *)
FUNCTION_BLOCK DELAY
    (*http://www.oscat.de/images/OSCATBasic/oscat_basic333_en.pdf#page=274*)
    stop := LIMIT(0,N,32) - 1;
    IF RST OR NOT init THEN
    	init := TRUE;
    	FOR i := 0 TO stop DO buf[i] := IN; END_FOR
    	OUT := IN;
    	i := 0;
    ELSIF stop < 0 THEN
    	OUT := IN;
    ELSE
    	OUT := buf[i];
    	buf[i] := IN;
    	i := INC1(i, N);
    END_IF

    (* revision history
    hm 1.10.2006		rev 1.1
    	corrected error IN buffer management

    hm 19.1.2007		rev 1.2
    	changed reset to load the value of IN instead of 0

    hm	27. oct. 2008	rev 1.3
    	improved performance

    hm	23. feb.2009	rev 1.4
    	corrected an index problem

    hm	23. mar. 2009	rev 1.5
    	corrected non standard write to input N

    *)
END_FUNCTION_BLOCK

(* ---- DELAY_4.st ---- *)
FUNCTION_BLOCK DELAY_4
    (*http://www.oscat.de/images/OSCATBasic/oscat_basic333_en.pdf#page=275*)
    OUT4 := OUT3;
    OUT3 := OUT2;
    OUT2 := OUT1;
    OUT1 := temp;
    temp := IN;

    (* revision history

    hm 19.1.2007	rev 1.1
    	added variable temp to add 1 delay  for q1

    *)
END_FUNCTION_BLOCK

(* ---- DRIVER_1.st ---- *)
FUNCTION_BLOCK DRIVER_1
    (*http://www.oscat.de/images/OSCATBasic/oscat_basic333_en.pdf#page=454*)
    IF off.Q THEN Q := FALSE; END_IF
    IF RST THEN
    	Q := FALSE;
    ELSIF SET THEN
    	Q := TRUE;
    ELSIF IN AND NOT edge_ THEN
    	IF TOGGLE_MODE THEN Q := NOT Q; ELSE Q := TRUE; END_IF
    END_IF
    edge_ := IN;
    IF TIMEOUT > t#0s THEN off(IN := Q, PT := TIMEOUT); END_IF

    (* revision history
    hm	2. jan 2008		rev 1.0
    	original version

    *)
END_FUNCTION_BLOCK

(* ---- DRIVER_4.st ---- *)
FUNCTION_BLOCK DRIVER_4
    (*http://www.oscat.de/images/OSCATBasic/oscat_basic333_en.pdf#page=454*)
    d0(SET:=SET, IN:=IN0, RST:=RST, TOGGLE_MODE:=TOGGLE_MODE, TIMEOUT:=TIMEOUT);
    d1(SET:=SET, IN:=IN1, RST:=RST, TOGGLE_MODE:=TOGGLE_MODE, TIMEOUT:=TIMEOUT);
    d2(SET:=SET, IN:=IN2, RST:=RST, TOGGLE_MODE:=TOGGLE_MODE, TIMEOUT:=TIMEOUT);
    d3(SET:=SET, IN:=IN3, RST:=RST, TOGGLE_MODE:=TOGGLE_MODE, TIMEOUT:=TIMEOUT);
    Q0 := d0.Q;
    Q1 := d1.Q;
    Q2 := d2.Q;
    Q3 := d3.Q;

    (* revision history
    hm	2. jan 2008		rev 1.0
    	original version

    *)
END_FUNCTION_BLOCK

(* ---- DRIVER_4C.st ---- *)
FUNCTION_BLOCK DRIVER_4C
    (*http://www.oscat.de/images/OSCATBasic/oscat_basic333_en.pdf#page=455*)
    IF RST OR off.Q THEN
    	SN := 0;
    ELSIF IN AND NOT edge_ THEN
    	SN := SN + 1;
    	IF SN > 7 OR SX[SN] = 0 THEN SN := 0; END_IF
    END_IF
    edge_ := IN;
    IF SN > 0 THEN
    	Q0 := SX[SN].0;
    	Q1 := SX[SN].1;
    	Q2 := SX[SN].2;
    	Q3 := SX[SN].3;
    ELSE
    	Q0 := FALSE;
    	Q1 := FALSE;
    	Q2 := FALSE;
    	Q3 := FALSE;
    END_IF

    (* maximaum TIMEOUT *)
    IF TIMEOUT > t#0s THEN off(IN := SN > 0, PT := TIMEOUT); END_IF

    (* revision history
    hm	23. mar. 2009	rev 1.0
    	original version

    *)
END_FUNCTION_BLOCK

(* ---- DT_SIMU.st ---- *)
FUNCTION_BLOCK DT_SIMU
    (*http://www.oscat.de/images/OSCATBasic/oscat_basic333_en.pdf#page=338*)
    (* read system timer *)
    tx := T_PLC_MS();
    tc := REAL_TO_UDINT(UDINT_TO_REAL(tx - last) * SPEED);

    IF NOT init THEN
    	init := TRUE;
    	DTS := START;
    	tc := 0;
    	last := tx;
    ELSIF SPEED = 0.0 THEN
    	DTS := UDINT_TO_DT(DT_TO_UDINT(DTS) + 1);
    ELSIF tc >= 1000 THEN
    	td := (tc / 1000) * 1000;
    	DTS := DTS + UDINT_TO_TIME(td);
    	last := last + REAL_TO_UDINT(UDINT_TO_REAL(td) / SPEED);
    END_IF

    (* revision history
    hm	11. sep. 2008	rev 1.0
    	original version

    hm	16. nov	2008	rev 1.1
    	added type conversions for compatibility reasons

    hm	8.	mar. 2009	rev 1.2
    	added increment by cycle mode

    *)

END_FUNCTION_BLOCK

(* ---- ENERGY.st ---- *)
FUNCTION_BLOCK ENERGY
    (*http://www.oscat.de/images/OSCATBasic/oscat_basic333_en.pdf#page=361*)
    YJ := J + WH * 3600.0 + C * 4.1868;
    YC := YJ * 0.238845896627496;
    YWH := YJ * 2.7777777778E-004;

    (*
    Arbeit, Energie, Joule* J 1 J = 1 N · m = 1 W · s = (1/3,6) E–6 kW · h = 1 kg · m2/s2
    Wärmemenge Kilowattstunde kW · h 1 kW · h = 3,6 MJ = 860 kcal
    Elektronvolt eV 1 eV = 160,218 92 E–21 J
    Erg erg 1 erg = 1E–7 J
    Kalorie calorie 1 calalorie = 4,1868 J = 1,163 E–3 W · h
    Therm therm 1 therm = 105,50 · 106 J
    *)

    (* revision history

    hm	27. mar. 2007	rev 1.0
    	original version

    hm	11. mar. 2009	rev 1.1
    	improved code

    hm 16. jan 2010	rev 1.2
    	avoid the string cal in comments for codesys import bug

    *)
END_FUNCTION_BLOCK

(* ---- ESR_COLLECT.st ---- *)
FUNCTION_BLOCK ESR_COLLECT
    (*http://www.oscat.de/images/OSCATBasic/oscat_basic333_en.pdf#page=33*)
    IF RST OR cnt < 0 THEN
    	POS := -1;
    ELSE
    	FOR cnt := 0 TO max_in DO
    	IF ESR_0[cnt].TYP > 0 THEN POS := INC1(POS, max_out); ESR_OUT[POS] := ESR_0[cnt]; END_IF
    	IF ESR_1[cnt].TYP > 0 THEN POS := INC1(POS, max_out); ESR_OUT[POS] := ESR_1[cnt]; END_IF
    	IF ESR_2[cnt].TYP > 0 THEN POS := INC1(POS, max_out); ESR_OUT[POS] := ESR_2[cnt]; END_IF
    	IF ESR_3[cnt].TYP > 0 THEN POS := INC1(POS, max_out); ESR_OUT[POS] := ESR_3[cnt]; END_IF
    	IF ESR_4[cnt].TYP > 0 THEN POS := INC1(POS, max_out); ESR_OUT[POS] := ESR_4[cnt]; END_IF
    	IF ESR_5[cnt].TYP > 0 THEN POS := INC1(POS, max_out); ESR_OUT[POS] := ESR_5[cnt]; END_IF
    	IF ESR_6[cnt].TYP > 0 THEN POS := INC1(POS, max_out); ESR_OUT[POS] := ESR_6[cnt]; END_IF
    	IF ESR_7[cnt].TYP > 0 THEN POS := INC1(POS, max_out); ESR_OUT[POS] := ESR_7[cnt]; END_IF
       END_FOR
    END_IF

    (* revision history
    hm	26.jan 2007	rev 1.0
    	original version

    hm	8. dec 2007	rev 1.1
    	added reset input

    ks	27. oct. 2008	rev 1.2
    	optimized code for performance

    ks	12. nov. 2009	rev 1.3
    	output POS was not pointing to last value

    hm	1. dec. 2009	rev 1.4
    	changed POS to be I/O
    	reduced output array size to 32 elements
    *)
END_FUNCTION_BLOCK

(* ---- ESR_MON_B8.st ---- *)
FUNCTION_BLOCK ESR_MON_B8
    (*http://www.oscat.de/images/OSCATBasic/oscat_basic333_en.pdf#page=35*)
    (* read system timer *)
    tx := UDINT_TO_TIME(T_PLC_MS());

    ESR_FLAG := FALSE;
    ESR_OUT[3].TYP := 0;
    ESR_OUT[2].TYP := 0;
    ESR_OUT[1].TYP := 0;
    ESR_OUT[0].TYP := 0;
    cnt := 0;

    (* check if inputs have chaged and fill buffer *)
    IF S0 <> x0 THEN
    	ESR_OUT[cnt].TYP := 10;
        ESR_OUT[cnt].TYP.0 := S0;
    	ESR_OUT[cnt].ADRESS := A0;
    	ESR_OUT[cnt].DS := DT_IN;
    	ESR_OUT[cnt].TS := tx;
    	x0 := S0;
    	cnt := cnt + 1;
    	ESR_FLAG := TRUE;
    END_IF
    IF S1 <> x1 THEN
    	ESR_OUT[cnt].TYP := 10;
        ESR_OUT[cnt].TYP.0 := S1;
    	ESR_OUT[cnt].ADRESS := A1;
    	ESR_OUT[cnt].DS := DT_IN;
    	ESR_OUT[cnt].TS := tx;
    	x1 := S1;
    	cnt := cnt + 1;
    	ESR_FLAG := TRUE;
    END_IF
    IF S2 <> x2 THEN
    	ESR_OUT[cnt].TYP := 10;
        ESR_OUT[cnt].TYP.0 := S2;
    	ESR_OUT[cnt].ADRESS := A2;
    	ESR_OUT[cnt].DS := DT_IN;
    	ESR_OUT[cnt].TS := tx;
    	x2 := S2;
    	cnt := cnt + 1;
    	ESR_FLAG := TRUE;
    END_IF
    IF S3 <> x3 THEN
    	ESR_OUT[cnt].TYP := 10;
        ESR_OUT[cnt].TYP.0 := S3;
    	ESR_OUT[cnt].ADRESS := A3;
    	ESR_OUT[cnt].DS := DT_IN;
    	ESR_OUT[cnt].TS := tx;
    	x3 := S3;
    	cnt := cnt + 1;
    	ESR_FLAG := TRUE;
    END_IF
    IF S4 <> x4 AND cnt < 4 THEN
    	ESR_OUT[cnt].TYP := 10;
        ESR_OUT[cnt].TYP.0 := S4;
    	ESR_OUT[cnt].ADRESS := A4;
    	ESR_OUT[cnt].DS := DT_IN;
    	ESR_OUT[cnt].TS := tx;
    	x4 := S4;
    	cnt := cnt + 1;
    	ESR_FLAG := TRUE;
    END_IF
    IF S5 <> x5  AND cnt < 4 THEN
    	ESR_OUT[cnt].TYP := 10;
        ESR_OUT[cnt].TYP.0 := S5;
    	ESR_OUT[cnt].ADRESS := A5;
    	ESR_OUT[cnt].DS := DT_IN;
    	ESR_OUT[cnt].TS := tx;
    	x5 := S5;
    	cnt := cnt + 1;
    	ESR_FLAG := TRUE;
    END_IF
    IF S6 <> x6  AND cnt < 4 THEN
    	ESR_OUT[cnt].TYP := 10;
        ESR_OUT[cnt].TYP.0 := S6;
    	ESR_OUT[cnt].ADRESS := A6;
    	ESR_OUT[cnt].DS := DT_IN;
    	ESR_OUT[cnt].TS := tx;
    	x6 := S6;
    	cnt := cnt + 1;
    	ESR_FLAG := TRUE;
    END_IF
    IF S7 <> x7  AND cnt < 4 THEN
    	ESR_OUT[cnt].TYP := 10;
        ESR_OUT[cnt].TYP.0 := S7;
    	ESR_OUT[cnt].ADRESS := A7;
    	ESR_OUT[cnt].DS := DT_IN;
    	ESR_OUT[cnt].TS := tx;
    	x7 := S7;
    	cnt := cnt + 1;
    	ESR_FLAG := TRUE;
    END_IF

    (* revision history
    hm	26. jan 2007	rev 1.0
    	original version

    hm	17. sep 2007	rev 1.1
    	replaced time() with T_PLC_MS() for compatibility reasons

    hm	22. oct. 2008	rev 1.2
    	optimized code

    hm	1.dec. 2009	rev 1.3
    	changed ESR_OUT to be I/O

    *)
END_FUNCTION_BLOCK

(* ---- ESR_MON_R4.st ---- *)
FUNCTION_BLOCK ESR_MON_R4
    (*http://www.oscat.de/images/OSCATBasic/oscat_basic333_en.pdf#page=35*)
    (* read system timer *)
    tx := UDINT_TO_TIME(T_PLC_MS());
    p0 ACCESS ADR(R0);
    p1 ACCESS ADR(R1);
    p2 ACCESS ADR(R2);
    p3 ACCESS ADR(R3);

    ESR_FLAG := FALSE;
    ESR_OUT[3].TYP := 0;
    ESR_OUT[2].TYP := 0;
    ESR_OUT[1].TYP := 0;
    ESR_OUT[0].TYP := 0;
    cnt := 0;

    (* check if inputs have chaged and fill buffer *)
    IF DIFFER(R0,  x0, S0) THEN
    	ESR_OUT[cnt].TYP := 20;
    	ESR_OUT[cnt].ADRESS := A0;
    	ESR_OUT[cnt].DS := DT_IN;
    	ESR_OUT[cnt].TS := tx;
    	ESR_OUT[cnt].DATA[0] := BYTE_OF_DWORD(p0,0);
    	ESR_OUT[cnt].DATA[1] := BYTE_OF_DWORD(p0,1);
    	ESR_OUT[cnt].DATA[2] := BYTE_OF_DWORD(p0,2);
    	ESR_OUT[cnt].DATA[3] := BYTE_OF_DWORD(p0,3);
    	x0 := R0;
    	cnt := cnt + 1;
    	ESR_FLAG := TRUE;
    END_IF
    IF DIFFER(R1,  x1, S1) THEN
    	ESR_OUT[cnt].TYP := 20;
    	ESR_OUT[cnt].ADRESS := A1;
    	ESR_OUT[cnt].DS := DT_IN;
    	ESR_OUT[cnt].TS := tx;
    	ESR_OUT[cnt].DATA[0] := BYTE_OF_DWORD(p1,0);
    	ESR_OUT[cnt].DATA[1] := BYTE_OF_DWORD(p1,1);
    	ESR_OUT[cnt].DATA[2] := BYTE_OF_DWORD(p1,2);
    	ESR_OUT[cnt].DATA[3] := BYTE_OF_DWORD(p1,3);
    	x1 := R1;
    	cnt := cnt + 1;
    	ESR_FLAG := TRUE;
    END_IF
    IF DIFFER(R2,  x2, S2) THEN
    	ESR_OUT[cnt].TYP := 20;
    	ESR_OUT[cnt].ADRESS := A2;
    	ESR_OUT[cnt].DS := DT_IN;
    	ESR_OUT[cnt].TS := tx;
    	ESR_OUT[cnt].DATA[0] := BYTE_OF_DWORD(p2,0);
    	ESR_OUT[cnt].DATA[1] := BYTE_OF_DWORD(p2,1);
    	ESR_OUT[cnt].DATA[2] := BYTE_OF_DWORD(p2,2);
    	ESR_OUT[cnt].DATA[3] := BYTE_OF_DWORD(p2,3);
    	x2 := R2;
    	cnt := cnt + 1;
    	ESR_FLAG := TRUE;
    END_IF
    IF DIFFER(R3,  x3, S3) THEN
    	ESR_OUT[cnt].TYP := 20;
    	ESR_OUT[cnt].ADRESS := A3;
    	ESR_OUT[cnt].DS := DT_IN;
    	ESR_OUT[cnt].TS := tx;
    	ESR_OUT[cnt].DATA[0] := BYTE_OF_DWORD(p3,0);
    	ESR_OUT[cnt].DATA[1] := BYTE_OF_DWORD(p3,1);
    	ESR_OUT[cnt].DATA[2] := BYTE_OF_DWORD(p3,2);
    	ESR_OUT[cnt].DATA[3] := BYTE_OF_DWORD(p3,3);
    	x3 := R3;
    	cnt := cnt + 1;
    	ESR_FLAG := TRUE;
    END_IF

    (* revision history
    hm	26. jan 2007	rev 1.0
    	original version

    hm	17. sep. 2007		rev 1.1
    	replaced time() with T_PLC_MS() for compatibility reasons

    hm	8. dec. 2007		rev 1.2
    	corrected an error while esr typ would not be set

    hm	16. mar. 2008		rev 1.3
    	deleted wrong conversion real_to_dword

    hm	1. dec 2009		rev 1.4
    	changed ESR_OUT to be I/O

    *)

END_FUNCTION_BLOCK

(* ---- ESR_MON_X8.st ---- *)
FUNCTION_BLOCK ESR_MON_X8
    (*http://www.oscat.de/images/OSCATBasic/oscat_basic333_en.pdf#page=36*)
    (* read system timer *)
    tx := UDINT_TO_TIME(T_PLC_MS());

    ESR_FLAG := FALSE;
    ESR_OUT[3].TYP := 0;
    ESR_OUT[2].TYP := 0;
    ESR_OUT[1].TYP := 0;
    ESR_OUT[0].TYP := 0;
    cnt := 0;

    (* check if inputs have chaged and fill buffer *)
    IF S0 <> x0 AND ((S0 < 100) OR (S0 > 99 AND S0 < 200 AND MODE >= 2) OR (S0 > 199 AND MODE = 3)) THEN
    	STATUS_TO_ESR(S0, A0, DT_IN, tx,ESR_OUT[cnt]);
    	x0 := S0;
    	cnt := cnt + 1;
    	ESR_FLAG := TRUE;
    END_IF
    IF S1 <> x1 AND ((S1 < 100) OR (S1 > 99 AND S1 < 200 AND MODE >= 2) OR (S1 > 199 AND MODE = 3)) THEN
    	STATUS_TO_ESR(S1, A1, DT_IN, tx,ESR_OUT[cnt]);
    	x1 := S1;
    	cnt := cnt + 1;
    	ESR_FLAG := TRUE;
    END_IF
    IF S2 <> x2 AND ((S2 < 100) OR (S2 > 99 AND S2 < 200 AND MODE >= 2) OR (S2 > 199 AND MODE = 3)) THEN
    	STATUS_TO_ESR(S2, A2, DT_IN, tx,ESR_OUT[cnt]);
    	x2 := S2;
    	cnt := cnt + 1;
    	ESR_FLAG := TRUE;
    END_IF
    IF S3 <> x3 AND ((S3 < 100) OR (S3 > 99 AND S3 < 200 AND MODE >= 2) OR (S3 > 199 AND MODE = 3)) THEN
    	STATUS_TO_ESR(S3, A3, DT_IN, tx,ESR_OUT[cnt]);
    	x3 := S3;
    	cnt := cnt + 1;
    	ESR_FLAG := TRUE;
    END_IF
    IF cnt < 4 AND S4 <> x4 AND ((S4 < 100) OR (S4 > 99 AND S4 < 200 AND MODE >= 2) OR (S4 > 199 AND MODE = 3)) THEN
    	STATUS_TO_ESR(S4, A4, DT_IN, tx,ESR_OUT[cnt]);
    	x4 := S4;
    	cnt := cnt + 1;
    	ESR_FLAG := TRUE;
    END_IF
    IF cnt < 4 AND S5 <> x5 AND ((S5 < 100) OR (S5 > 99 AND S5 < 200 AND MODE >= 2) OR (S5 > 199 AND MODE = 3)) THEN
    	STATUS_TO_ESR(S5, A5, DT_IN, tx,ESR_OUT[cnt]);
    	x5 := S5;
    	cnt := cnt + 1;
    	ESR_FLAG := TRUE;
    END_IF
    IF cnt < 4 AND S6 <> x6 AND ((S6 < 100) OR (S6 > 99 AND S6 < 200 AND MODE >= 2) OR (S6 > 199 AND MODE = 3)) THEN
    	STATUS_TO_ESR(S6, A6, DT_IN, tx,ESR_OUT[cnt]);
    	x6 := S6;
    	cnt := cnt + 1;
    	ESR_FLAG := TRUE;
    END_IF
    IF cnt < 4 AND S7 <> x7 AND ((S7 < 100) OR (S7 > 99 AND S7 < 200 AND MODE >= 2) OR (S7 > 199 AND MODE = 3)) THEN
    	STATUS_TO_ESR(S7, A7, DT_IN, tx,ESR_OUT[cnt]);
    	x7 := S7;
    	cnt := cnt + 1;
    	ESR_FLAG := TRUE;
    END_IF

    (* revision history
    hm	26. jan 2007		rev 1.0
    	original version

    hm	17. sep 2007	rev 1.1
    	replaced time() with T_PLC_MS() for compatibility reasons

    hm	1. dec. 2009	rev 1.2
    	changed ESR_OUT to be I/O

    *)
END_FUNCTION_BLOCK

(* ---- EVENTS.st ---- *)
FUNCTION_BLOCK EVENTS
    (*http://www.oscat.de/images/OSCATBasic/oscat_basic333_en.pdf#page=122*)
    (* for performance reasons only activate once a day *)
    IF last_active <> DATE_IN THEN
    	last_active := DATE_IN;
    	y_int := FALSE;
    	name_int := '';
    	day_in := DAY_OF_DATE(DATE_IN);
    	cyr := YEAR_OF_DATE(DATE_IN);

    	(* search list for events *)
    	FOR i := 0 TO size DO
    		check := ELIST[i];
    		lday := DAY_OF_DATE(SET_DATE(cyr,check.MONTH, check.DAY));
    		IF day_in >= lday AND day_in <= lday + check.USE - 1 THEN
    			y_int := TRUE;
    			name_int := check.NAME;
    			EXIT;
    		END_IF
    	END_FOR
    END_IF

    IF ENA THEN
    	Y := y_int;
    	NAME := name_int;
    ELSE
    	Y := FALSE;
    	NAME := '';
    END_IF

    (* revision history
    hm  18. jan. 2011	rev 1.0
    	new module

    *)

END_FUNCTION_BLOCK
